// Library/Functions/Swap/SwapIecDate
FUNCTION SwapIecDate : IEC_DATE
// ------------------------------------------------------------------------- 
//  SRCI Robot Library                                                
// ------------------------------------------------------------------------- 
//                                                                           
//  Object:      SwapIecDate                                       
//  Author:      Thorsten Brach                                                
//  Date:        2024-06-09
//
//  Description:                                              
//   
//                                                                           
//  Copyright: 
//    (C) 2024 Thorsten Brach. All rights reserved                                                                                                                                            
//             Licensed under the MIT License.
//                                                                           
//  Disclaimer:                                                                           
//    This project is provided without any guarantee and can be used for   
//    private and commercial purposes. Any use is at the user’s 
//    own risk and responsibility.
//
// -------------------------------------------------------------------------
VAR_INPUT
  /// Value to swap
  Value : IEC_DATE;
END_VAR

SwapBytes(ADR(Value),SIZEOF(Value));

SwapIecDate := Value;

END_FUNCTION

// Library/Functions/Swap/SwapIecTime
FUNCTION SwapIecTime : TOD
// ------------------------------------------------------------------------- 
//  SRCI Robot Library                                                
// ------------------------------------------------------------------------- 
//                                                                           
//  Object:      SwapTime                                       
//  Author:      Thorsten Brach                                                
//  Date:        2024-06-01
//
//  Description:                                              
//   
//                                                                           
//  Copyright: 
//    (C) 2024 Thorsten Brach. All rights reserved                                                                                                                                            
//             Licensed under the MIT License.
//                                                                           
//  Disclaimer:                                                                           
//    This project is provided without any guarantee and can be used for   
//    private and commercial purposes. Any use is at the user’s 
//    own risk and responsibility.
//
// -------------------------------------------------------------------------
VAR_INPUT
  /// Value
  Value : TOD;
END_VAR

SwapBytes(ADR(Value),SIZEOF(Value));

SwapIecTime := Value;

END_FUNCTION

// Library/Functions/Swap/SwapInt
FUNCTION SwapInt : INT
// ------------------------------------------------------------------------- 
//  SRCI Robot Library                                                
// ------------------------------------------------------------------------- 
//                                                                           
//  Object:      SwapInt                                       
//  Author:      Thorsten Brach                                                
//  Date:        2024-06-01
//
//  Description:                                              
//   
//                                                                           
//  Copyright: 
//    (C) 2024 Thorsten Brach. All rights reserved                                                                                                                                            
//             Licensed under the MIT License.
//                                                                           
//  Disclaimer:                                                                           
//    This project is provided without any guarantee and can be used for   
//    private and commercial purposes. Any use is at the user’s 
//    own risk and responsibility.
//
// -------------------------------------------------------------------------
VAR_INPUT
  /// Value to swap
  Value : INT;
END_VAR

SwapBytes(ADR(Value),SIZEOF(Value));

SwapInt := Value;

END_FUNCTION

// Library/Functions/Swap/SwapReal
FUNCTION SwapReal : REAL
// ------------------------------------------------------------------------- 
//  SRCI Robot Library                                                
// ------------------------------------------------------------------------- 
//                                                                           
//  Object:      SwapReal                                       
//  Author:      Thorsten Brach                                                
//  Date:        2024-06-01
//
//  Description:                                              
//   
//                                                                           
//  Copyright: 
//    (C) 2024 Thorsten Brach. All rights reserved                                                                                                                                            
//             Licensed under the MIT License.
//                                                                           
//  Disclaimer:                                                                           
//    This project is provided without any guarantee and can be used for   
//    private and commercial purposes. Any use is at the user’s 
//    own risk and responsibility.
//
// -------------------------------------------------------------------------
VAR_INPUT
  /// Value
  Value : REAL;
END_VAR

SwapBytes(ADR(Value),SIZEOF(Value));

SwapReal := Value;

END_FUNCTION

// Library/Functions/Swap/SwapUdint
FUNCTION SwapUdint : UDINT
// ------------------------------------------------------------------------- 
//  SRCI Robot Library                                                
// ------------------------------------------------------------------------- 
//                                                                           
//  Object:      SwapUdint                                       
//  Author:      Thorsten Brach                                                
//  Date:        2024-06-01
//
//  Description:                                              
//   
//                                                                           
//  Copyright: 
//    (C) 2024 Thorsten Brach. All rights reserved                                                                                                                                            
//             Licensed under the MIT License.
//                                                                           
//  Disclaimer:                                                                           
//    This project is provided without any guarantee and can be used for   
//    private and commercial purposes. Any use is at the user’s 
//    own risk and responsibility.
//
// -------------------------------------------------------------------------
VAR_INPUT
  /// Value
  Value : UDINT;
END_VAR

SwapBytes(ADR(Value),SIZEOF(Value));

SwapUdint := Value;

END_FUNCTION

// Library/Functions/Swap/SwapUint
FUNCTION SwapUint : UINT
// ------------------------------------------------------------------------- 
//  SRCI Robot Library                                                
// ------------------------------------------------------------------------- 
//                                                                           
//  Object:      SwapUint                                       
//  Author:      Thorsten Brach                                                
//  Date:        2024-06-01
//
//  Description:                                              
//   
//                                                                           
//  Copyright: 
//    (C) 2024 Thorsten Brach. All rights reserved                                                                                                                                            
//             Licensed under the MIT License.
//                                                                           
//  Disclaimer:                                                                           
//    This project is provided without any guarantee and can be used for   
//    private and commercial purposes. Any use is at the user’s 
//    own risk and responsibility.
//
// -------------------------------------------------------------------------
VAR_INPUT
  /// Value to swap
  Value : UINT;
END_VAR

SwapBytes(ADR(Value),SIZEOF(Value));

SwapUint := Value;

END_FUNCTION

// Library/Interfaces/IMessageLogger
INTERFACE IMessageLogger

METHOD PUBLIC AddMessageLog
VAR_INPUT
  /// Message to add to the log
  MessageLog : AlarmMessage;
END_VAR
END_METHOD

METHOD PUBLIC AddSystemLog
VAR_INPUT
  /// System messafe to add to the log
  SystemLog : STRING(RobotLibraryParameter.MESSAGE_TEXT_LEN);
END_VAR
END_METHOD

END_INTERFACE

// Library/Interfaces/IRobotLibraryCommandFB
INTERFACE IRobotLibraryCommandFB

METHOD PUBLIC CallBack : DINT
VAR_INPUT
  /// Response data
  RspData : AxesGroupAcyclicAcrEntryRspBuffer;  
END_VAR
END_METHOD

PROPERTY CommandData : RobotLibrarySendDataFB
GET
END_GET
SET
END_SET
END_PROPERTY

END_INTERFACE

// Library/POUs/_internal/Send/RobotLibrarySendDataFB
{attribute 'pack_mode' := '1'} 
FUNCTION_BLOCK RobotLibrarySendDataFB extends RobotLibrarySendDataBaseFB
// ------------------------------------------------------------------------- 
//  SRCI Robot Library                                                
// ------------------------------------------------------------------------- 
//                                                                           
//  Object:      RobotLibrarySendDataFB                                      
//  Author:      Thorsten Brach                                                
//  Date:        2024-06-01
//
//  Description:                                              
//    
//                                                                           
//  Copyright: 
//    (C) 2024 Thorsten Brach. All rights reserved                                                                                                                                            
//             Licensed under the MIT License.
//                                                                           
//  Disclaimer:                                                                           
//    This project is provided without any guarantee and can be used for   
//    private and commercial purposes. Any use is at the user’s 
//    own risk and responsibility.
//
// -------------------------------------------------------------------------
VAR_INPUT
  /// Payload
  Payload     : POINTER TO BYTE;
  /// Size of the Payload array
  PayLoadSize : UDINT;
END_VAR

/// Resets the payload buffer, the payload pointer and the payload length
METHOD Reset
VAR_INPUT
END_VAR
SUPER^.Reset();

// Reset payload buffer
SysDepMemSet(pDest := Payload, Value := 0 , DataLen := PayLoadSize);
END_METHOD

METHOD SetLifeSignFooter
VAR_INPUT
  /// Life sign value
  LifeSign : BYTE;
END_VAR

VAR
  /// temporary 
  pLifeSign : POINTER TO BYTE;
END_VAR
pLifeSign := Payload + PayLoadSize -1;

pLifeSign^ := LifeSign;
END_METHOD

METHOD UpdatePointer
VAR_INPUT
END_VAR
pPayload := Payload;
END_METHOD

END_FUNCTION_BLOCK

// Library/POUs/_internal/Send/RobotLibrarySendDataBaseFB
{attribute 'pack_mode' := '1'} 
FUNCTION_BLOCK RobotLibrarySendDataBaseFB
// ------------------------------------------------------------------------- 
//  SRCI Robot Library                                                
// ------------------------------------------------------------------------- 
//                                                                           
//  Object:      RobotLibrarySendDataFB                                      
//  Author:      Thorsten Brach                                                
//  Date:        2024-06-01
//
//  Description:                                              
//    
//                                                                           
//  Copyright: 
//    (C) 2024 Thorsten Brach. All rights reserved                                                                                                                                            
//             Licensed under the MIT License.
//                                                                           
//  Disclaimer:                                                                           
//    This project is provided without any guarantee and can be used for   
//    private and commercial purposes. Any use is at the user’s 
//    own risk and responsibility.
//
// -------------------------------------------------------------------------
VAR_INPUT
  /// Payload length
  PayloadLen : UDINT;
  /// Payload pointer
  PayloadPtr : UDINT;
END_VAR


VAR
  /// internal pointer to payload 
  pPayload : POINTER TO BYTE;
END_VAR

/// Adds a ArmConfigParameter to the payload buffer, increase the payload pointer and returns the payload lenght
METHOD AddArmConfig : UDINT
VAR_INPUT
  /// Value to add
  Value : ArmConfigParameter;
END_VAR

VAR
  /// temporary Byte
 _tmpByte : BYTE;
END_VAR
// Table 6-274: "ConfigMode" on "Command Management Layer"
// --------------------------
// --------------------------
// Byte 00 : Bit 00  - Shoulder
//         : Bit 01  - Shoulder
//         : Bit 02  - Shoulder
//         : Bit 03  - Shoulder
//         : Bit 04  - Elbow
//         : Bit 05  - Elbow
//         : Bit 06  - Elbow
//         : Bit 07  - Elbow
// Byte 01 : Bit 00  - Wrist
//         : Bit 01  - Wrist
//         : Bit 02  - Wrist
//         : Bit 03  - Wrist
//         : Bit 04  - Reserve
//         : Bit 05  - Reserve
//         : Bit 06  - Reserve
//         : Bit 07  - Reserve
_tmpByte.0 := Value.Shoulder = ArmConfigShoulder.BACK;
_tmpByte.1 := Value.Elbow    = ArmConfigElbow.DOWN;
_tmpByte.2 := Value.Wrist    = ArmConfigWrist.FLIP;

AddByte(_tmpByte);
AddByte(0);

AddArmConfig := PayloadLen;
END_METHOD

/// Adds a BOOL to the payload buffer, increase the payload pointer and returns the payload lenght
METHOD AddBool : UDINT
VAR_INPUT
  /// Value to add
  Value : BOOL;
END_VAR

VAR
  /// temporary byte
 _tmpByte : BYTE := 0;
END_VAR
// update internal pointer
UpdatePointer();

// check pointer is valid ? 
IF (pPayload = RobotLibraryConstants.NULL_POINTER)
THEN
  RETURN;
END_IF


_tmpByte.0 := Value;
// copy data 
SysDepMemCpy(pDest := pPayload + PayloadPtr, pSrc := ADR(_tmpByte), DataLen := SIZEOF(_tmpByte));
// inc payload pointer 
PayloadPtr := PayloadPtr + SIZEOF(_tmpByte);
// return payload len
AddBool := PayloadLen := PayloadPtr;
END_METHOD

/// Adds a BYTE to the payload buffer, increase the payload pointer and returns the payload lenght
METHOD AddByte : UDINT
VAR_INPUT
  /// Value to add
  Value : BYTE;
END_VAR
// update internal pointer
UpdatePointer();

// check pointer is valid ? 
IF (pPayload = RobotLibraryConstants.NULL_POINTER)
THEN
  RETURN;
END_IF


Value := Value;
// copy data 
SysDepMemCpy( pDest := pPayload + PayloadPtr, pSrc := ADR(Value), DataLen := SIZEOF(Value));
// inc payload pointer 
PayloadPtr := PayloadPtr + SIZEOF(Value);
// return payload len
AddByte := PayloadLen := PayloadPtr;
END_METHOD

/// Adds a DataBlock to the payload buffer, increase the payload pointer and returns the payload lenght
METHOD AddDataBlock : UDINT
VAR_INPUT
  /// Value to add
  pValue : POINTER TO BYTE;
  /// Size of data block
  Size   : UDINT;
END_VAR
// update internal pointer
UpdatePointer();

// check pointer is valid ? 
IF (pPayload = RobotLibraryConstants.NULL_POINTER)
THEN
  RETURN;
END_IF


IF (pValue = 0) OR (Size = 0 )
THEN
  RETURN;
END_IF

// copy data 
SysDepMemCpy( pDest := pPayload + PayloadPtr, pSrc := pValue, DataLen := Size);
// inc payload pointer 
PayloadPtr := PayloadPtr + Size;
// return payload len
AddDataBlock := PayloadLen := PayloadPtr;
END_METHOD

/// Adds a DataInSync to the payload buffer, increase the payload pointer and returns the payload lenght
METHOD AddDataEnableSync : UDINT
VAR_INPUT
  /// Value to add
  Value : DataEnableSync;
END_VAR

VAR
  /// temporary Byte
 _tmpByte : BYTE;
END_VAR
Value := Value;

_tmpByte.0 := Value.EnableSyncTool;
_tmpByte.1 := Value.EnableSyncFrame;
_tmpByte.2 := Value.EnableSyncLoad;
_tmpByte.3 := Value.EnableSyncWorkArea;
_tmpByte.4 := Value.EnableSyncSWLimits;
_tmpByte.5 := Value.EnableSyncDefaultDynamics;
_tmpByte.6 := Value.EnableSyncReferenceDynamics;


AddByte(_tmpByte);

AddDataEnableSync := PayloadLen;
END_METHOD

/// Adds a DataInSync to the payload buffer, increase the payload pointer and returns the payload lenght
METHOD AddDataInSync : UDINT
VAR_INPUT
  /// Value to add
  Value : DataInSync;
END_VAR

VAR
  /// temporary Byte
 _tmpByte : BYTE;
END_VAR
Value := Value;

_tmpByte.0 := Value.ToolsInSync;
_tmpByte.1 := Value.FramesInSync;
_tmpByte.2 := Value.LoadsInSync;
_tmpByte.3 := Value.WorkAreasInSync;
_tmpByte.4 := Value.SoftwareLimitsInSync;
_tmpByte.5 := Value.DefaultDynamicsInSync;
_tmpByte.6 := Value.ReferenceDynamicsInSync;
_tmpByte.7 := FALSE;

AddByte(_tmpByte);

AddDataInSync := PayloadLen;
END_METHOD

/// Adds a DWORD to the payload buffer , increase the payload pointer and returns the payload lenght
METHOD AddDword : UDINT
VAR_INPUT
  /// Value to add
  Value : DWORD;
END_VAR
// update internal pointer
UpdatePointer();

// check pointer is valid ? 
IF (pPayload = RobotLibraryConstants.NULL_POINTER)
THEN
  RETURN;
END_IF


// swap byte order
Value := SwapDword(Value);
// copy data 
SysDepMemCpy(pDest := pPayload + PayloadPtr, pSrc := ADR(Value), DataLen := SIZEOF(Value));
// inc data index 
PayloadPtr := PayloadPtr + SIZEOF(Value);
// return payload len
AddDword := PayloadLen := PayloadPtr;
END_METHOD

/// Adds two halfe BYTE to the payload buffer , increase the payload pointer and returns the payload lenght
METHOD AddHalfBytes : UDINT
VAR_INPUT
  /// Value to add
  HalfByteHi : BYTE;
  /// Value to add
  HalfByteLo : BYTE;
END_VAR

VAR
  /// internal value
 _value : BYTE;
END_VAR
// update internal pointer
UpdatePointer();

// check pointer is valid ? 
IF (pPayload = RobotLibraryConstants.NULL_POINTER)
THEN
  RETURN;
END_IF


_value := CombineHalfBytes( HalfByteHi := HalfByteHi, HalfByteLo := HalfByteLo);
// copy data 
SysDepMemCpy(pDest := pPayload + PayloadPtr, pSrc := ADR(_value), DataLen := SIZEOF(_value));
// inc payload pointer 
PayloadPtr := PayloadPtr + SIZEOF(_value);
// return payload len
AddHalfBytes := PayloadLen := PayloadPtr;
END_METHOD

/// Adds a IEC_DATE to the payload buffer, increase the payload pointer and returns the payload lenght
METHOD AddIecDate : UDINT
VAR_INPUT
  /// Value to add
  Value : IEC_DATE;
END_VAR
// update internal pointer
UpdatePointer();

// check pointer is valid ? 
IF (pPayload = RobotLibraryConstants.NULL_POINTER)
THEN
  RETURN;
END_IF


Value := SwapIecDate(Value);
// copy data 
SysDepMemCpy(pDest := pPayload + PayloadPtr, pSrc := ADR(Value), DataLen := SIZEOF(Value));
// inc payload pointer 
PayloadPtr := PayloadPtr + SIZEOF(Value);
// return payload len
AddIecDate := PayloadLen := PayloadPtr;
END_METHOD

/// Adds a IEC_TIME to the payload buffer, increase the payload pointer and returns the payload lenght
METHOD AddIecTime : UDINT
VAR_INPUT
  /// Value to add
  Value : IEC_TIME;
END_VAR
// update internal pointer
UpdatePointer();

// check pointer is valid ? 
IF (pPayload = RobotLibraryConstants.NULL_POINTER)
THEN
  RETURN;
END_IF


Value := SwapIecTime(Value);
// copy data 
SysDepMemCpy(pDest := pPayload + PayloadPtr, pSrc := ADR(Value), DataLen := SIZEOF(Value));
// inc payload pointer 
PayloadPtr := PayloadPtr + SIZEOF(Value);
// return payload len
AddIecTime := PayloadLen := PayloadPtr;
END_METHOD

/// Adds a INT to the payload buffer , increase the payload pointer and returns the payload lenght
METHOD AddInt : UDINT
VAR_INPUT
  /// Value to add
  Value : INT;
END_VAR
// update internal pointer
UpdatePointer();

// check pointer is valid ? 
IF (pPayload = RobotLibraryConstants.NULL_POINTER)
THEN
  RETURN;
END_IF


// swap byte order
Value := SwapInt(Value);
// copy data 
SysDepMemCpy(pDest := pPayload + PayloadPtr, pSrc := ADR(Value), DataLen := SIZEOF(Value));
// inc data index 
PayloadPtr := PayloadPtr + SIZEOF(Value);
// return payload len
AddInt := PayloadLen := PayloadPtr;
END_METHOD

/// Adds a REAL to the payload buffer , increase the payload pointer and returns the payload lenght
METHOD AddReal : UDINT
VAR_INPUT
  /// Value to add
  Value : REAL;
END_VAR
// update internal pointer
UpdatePointer();

// check pointer is valid ? 
IF (pPayload = RobotLibraryConstants.NULL_POINTER)
THEN
  RETURN;
END_IF


// swap byte order
Value := SwapReal(Value);
// copy data 
SysDepMemCpy(pDest := pPayload + PayloadPtr,pSrc := ADR(Value), DataLen := SIZEOF(Value));
// inc data index 
PayloadPtr := PayloadPtr + SIZEOF(Value);
// return payload len
AddReal := PayloadLen := PayloadPtr;
END_METHOD

/// Adds a SINT to the payload buffer, increase the payload pointer and returns the payload lenght
METHOD AddSint : UDINT
VAR_INPUT
  /// Value to add
  Value : SINT;
END_VAR
// update internal pointer
UpdatePointer();

// check pointer is valid ? 
IF (pPayload = RobotLibraryConstants.NULL_POINTER)
THEN
  RETURN;
END_IF


Value := Value;
// copy data 
SysDepMemCpy(pDest := pPayload + PayloadPtr, pSrc := ADR(Value), DataLen := SIZEOF(Value));
// inc payload pointer 
PayloadPtr := PayloadPtr + SIZEOF(Value);
// return payload len
AddSint := PayloadLen := PayloadPtr;
END_METHOD

/// Adds a String to the payload buffer, increase the payload pointer and returns the payload lenght
METHOD AddString : UDINT
VAR_INPUT
  /// Value to add
  Value : STRING(255);
END_VAR
// update internal pointer
UpdatePointer();

// check pointer is valid ? 
IF (pPayload = RobotLibraryConstants.NULL_POINTER)
THEN
  RETURN;
END_IF


IF ( LEN(Value) = 0 )
THEN
  RETURN;
END_IF

// copy data 
SysDepMemCpy(pDest := pPayload + PayloadPtr, pSrc := ADR(Value), DataLen := DINT_TO_UDINT(LEN(Value)));
// inc payload pointer 
PayloadPtr := PayloadPtr + DINT_TO_UDINT(LEN(Value));
// return payload len
AddString := PayloadLen := PayloadPtr;
END_METHOD

/// Adds a TIME to the payload buffer , increase the payload pointer and returns the payload lenght
METHOD AddTime : UDINT
VAR_INPUT
  /// Value to add
  Value : TOD;
END_VAR
// update internal pointer
UpdatePointer();

// check pointer is valid ? 
IF (pPayload = RobotLibraryConstants.NULL_POINTER)
THEN
  RETURN;
END_IF


// swap byte order
Value := SwapIecTime(Value);
// copy data 
SysDepMemCpy(pDest := pPayload + PayloadPtr, pSrc := ADR(Value), DataLen := SIZEOF(Value));
// inc data index 
PayloadPtr := PayloadPtr + SIZEOF(Value);
// return payload len
AddTime := PayloadLen := PayloadPtr;
END_METHOD

/// Adds a TurnNumber to the payload buffer, increase the payload pointer and returns the payload lenght
METHOD AddTurnNumber : UDINT
VAR_INPUT
  /// Value to add
  Value : TurnNumber;
END_VAR

VAR
  /// temporary Byte
 _tmpByte : BYTE;
END_VAR
Value := Value;

// ST-FIX F3: sign + magnitude (spec 5.5.4.4)
AddHalfBytes( HalfByteHi := TURN_TO_SIGN_MAGNITUDE(Turns := Value.J2Turns, Bits := 3), HalfByteLo := TURN_TO_SIGN_MAGNITUDE(Turns := Value.J1Turns, Bits := 3));
AddHalfBytes( HalfByteHi := TURN_TO_SIGN_MAGNITUDE(Turns := Value.J4Turns, Bits := 3), HalfByteLo := TURN_TO_SIGN_MAGNITUDE(Turns := Value.J3Turns, Bits := 3));
AddHalfBytes( HalfByteHi := TURN_TO_SIGN_MAGNITUDE(Turns := Value.J6Turns, Bits := 3), HalfByteLo := TURN_TO_SIGN_MAGNITUDE(Turns := Value.J5Turns, Bits := 3));
AddByte(TURN_TO_SIGN_MAGNITUDE(Turns := Value.E1Turns, Bits := 7));

AddTurnNumber := PayloadLen;
END_METHOD

/// Adds a UDINT to the payload buffer , increase the payload pointer and returns the payload lenght
METHOD AddUdint : UDINT
VAR_INPUT
  /// Value to add
  Value : UDINT;
END_VAR
// update internal pointer
UpdatePointer();

// check pointer is valid ? 
IF (pPayload = RobotLibraryConstants.NULL_POINTER)
THEN
  RETURN;
END_IF


// swap byte order
Value := SwapUdint(Value);
// copy data 
SysDepMemCpy(pDest := pPayload + PayloadPtr, pSrc := ADR(Value), DataLen := SIZEOF(Value));
// inc data index 
PayloadPtr := PayloadPtr + SIZEOF(Value);
// return payload len
AddUdint := PayloadLen := PayloadPtr;
END_METHOD

/// Adds a UINT to the payload buffer , increase the payload pointer and returns the payload lenght
METHOD AddUint : UDINT
VAR_INPUT
  /// Value to add
  Value : UINT;
END_VAR
// update internal pointer
UpdatePointer();

// check pointer is valid ? 
IF (pPayload = RobotLibraryConstants.NULL_POINTER)
THEN
  RETURN;
END_IF


// swap byte order
Value := SwapUint(Value);
// copy data 
SysDepMemCpy(pDest := pPayload + PayloadPtr, pSrc := ADR(Value), DataLen := SIZEOF(Value));
// inc data index 
PayloadPtr := PayloadPtr + SIZEOF(Value);
// return payload len
AddUint := PayloadLen := PayloadPtr;
END_METHOD

/// Adds a USINT to the payload buffer, increase the payload pointer and returns the payload lenght
METHOD AddUsint : UDINT
VAR_INPUT
  /// Value to add
  Value : USINT;
END_VAR
// update internal pointer
UpdatePointer();

// check pointer is valid ? 
IF (pPayload = RobotLibraryConstants.NULL_POINTER)
THEN
  RETURN;
END_IF


Value := Value;
// copy data 
SysDepMemCpy(pDest := pPayload + PayloadPtr, pSrc := ADR(Value), DataLen := SIZEOF(Value));
// inc payload pointer 
PayloadPtr := PayloadPtr + SIZEOF(Value);
// return payload len
AddUsint := PayloadLen := PayloadPtr;
END_METHOD

/// Resets the payload buffer, the payload pointer and the payload length
METHOD Reset
VAR_INPUT
END_VAR
PayloadLen := 0;
PayloadPtr := 0;
END_METHOD

METHOD UpdatePointer
VAR_INPUT
END_VAR
END_METHOD

END_FUNCTION_BLOCK

// Library/POUs/_internal/BaseFBs/RobotLibraryBaseEnableFB
FUNCTION_BLOCK RobotLibraryBaseEnableFB EXTENDS RobotLibraryBaseFB
// ------------------------------------------------------------------------- 
//  SRCI Robot Library                                                
// ------------------------------------------------------------------------- 
//                                                                           
//  Object:      RobotLibraryBaseFB                                       
//  Author:      Thorsten Brach                                                
//  Date:        2024-08-11
//
//  Description:                                              
//   
//                                                                           
//  Copyright: 
//    (C) 2024 Thorsten Brach. All rights reserved                                                                                                                                            
//             Licensed under the MIT License.
//                                                                           
//  Disclaimer:                                                                           
//    This project is provided without any guarantee and can be used for   
//    private and commercial purposes. Any use is at the user’s 
//    own risk and responsibility.
//
// -------------------------------------------------------------------------
VAR_INPUT
  /// Set TRUE to activate / Set False to deactivate
  Enable            : BOOL;
END_VAR

VAR_OUTPUT
  /// FB is being processed
  Busy              : BOOL;
  /// TRUE while function is active
  Enabled           : BOOL;
END_VAR

VAR
  /// Rising edge for enable
  {attribute 'hide'}
 _enable_R          : R_TRIG;
  /// Falling edge for enable
  {attribute 'hide'}
 _enable_F          : F_TRIG;
END_VAR

SUPER^(AxesGroup := AxesGroup);

// ST-FIX F135: "Enabled" is reset with the falling edge of "Enable" as soon as possible
// (spec 5.5.10 output status), also while the FB still sends the deactivation to the RC
IF ( NOT Enable )
THEN
  Enabled := FALSE;
END_IF

METHOD PROTECTED OnCall
VAR_IN_OUT
  /// Robot assignment of function
  AxesGroup : AxesGroup; 
END_VAR

VAR
  /// internal return value
 _retVal : DINT;
END_VAR

                  SUPER^.OnCall(AxesGroup := AxesGroup);

// building rising and falling edges
_enable_R( CLK := Enable);
_enable_F( CLK := Enable);


// Check command execution is allowed ?
IF ((     Enable                                 ) AND
    ( NOT AxesGroup.State.Initialized            ) AND
    ( NOT AxesGroup.State.Synchronized           ) AND
    (     MyType <> 'MC_ExchangeConfigurationFB' ) AND // is part of init sequence
    (     MyType <> 'MC_ReadMessagesFB'          ) AND // is part of init sequence
    (     MyType <> 'MC_ReadRobotDataFB'         ))    // is part of init sequence
THEN
  SetError( ErrorID := RobotLibraryErrorIdEnum.ERR_COMMANDS_NOT_ENABLED, Overwrite := TRUE );
  Error   := TRUE;
  Busy    := FALSE; 
END_IF


// On execution started
IF ( _enable_R.Q )
THEN
  // ST-FIX F23: a new enable ends a pending cancel / error clear of the previous enable
  _cancel := FALSE;
  _stepCancel := 0;
  _clearError := FALSE;
  _stepClearError := 0;
  // ST-FIX F78: an error of the previous enable that is still being cleared (falling edge, up
  // to 5 s) is cleared now - otherwise the block (start only without Error) consumes the
  // rising edge and the new enable is ignored (not sent, no Busy, no Error)
  IF ( Error ) AND ( ErrorID <> RobotLibraryErrorIdEnum.ERR_COMMANDS_NOT_ENABLED )
  THEN
    Reset();
  END_IF
  OnExecStart(AxesGroup := AxesGroup);
END_IF


// On execution cancel  
IF ( Busy ) AND ( _enable_F.Q ) 
THEN
  // set cancel flag
 _cancel := TRUE;
END_IF

IF ( _cancel )
THEN
  // call Cancel
 _retVal := OnExecCancel(AxesGroup := AxesGroup);
  
  // done or error ?
  IF ( _retVal <> RobotLibraryConstants.RUNNING )
  THEN
    // reset cancel flag
   _cancel := FALSE;
	END_IF
END_IF


// On execution error clear
IF ( Error ) AND ( _enable_F.Q )
THEN
  // set ClearError flag
 _clearError := TRUE;
END_IF

IF ( _clearError )
THEN
 _retVal := OnExecErrorClear(AxesGroup := AxesGroup); 

  // done or error ?
  IF ( _retVal <> RobotLibraryConstants.RUNNING )
  THEN
    // reset ClearError flag
   _clearError := FALSE;
	END_IF
END_IF
END_METHOD

METHOD Protected OnExecCancel : DINT
VAR_IN_OUT
  /// Robot assignment of function
  AxesGroup : AxesGroup; 
END_VAR
VAR
  /// internal return value 
 _retVal    : DINT;
END_VAR
OnExecCancel := Reset();

// Create log entry
CreateLogMessagePara1 ( Timestamp   := AxesGroup.State.SystemTime,
                        MessageType := MessageType.CMD,
                        Severity    := Severity.DEBUG,
                        MessageCode := 0,
                        MessageText := 'Execution of {1} cancled ',
                        Para1       := MyType);                 

// try to remove cmd
_retVal := AxesGroup.Acyclic.ActiveCommandRegister.RemoveCmd(_uniqueID);

IF (_retVal = RobotLibraryConstants.OK)
THEN
  // Create log entry
  CreateLogMessagePara1 ( Timestamp   := AxesGroup.State.SystemTime,
                          MessageType := MessageType.CMD,
                          Severity    := Severity.DEBUG,
                          MessageCode := 0,
                          MessageText := '{1} successfully removed from ACR',
                          Para1       := MyType);                 
ELSE
  // Create log entry
  CreateLogMessagePara1 ( Timestamp   := AxesGroup.State.SystemTime,
                          MessageType := MessageType.CMD,
                          Severity    := Severity.DEBUG,
                          MessageCode := 0,
                          MessageText := '{1} was not removed from ACR because execution was already in progress',
                          Para1       := MyType);                 
END_IF
END_METHOD

METHOD PROTECTED OnExecErrorClear : DINT
VAR_IN_OUT
  /// Robot assignment of function
  AxesGroup : AxesGroup; 
END_VAR
OnExecErrorClear := RobotLibraryConstants.RUNNING;

CASE _stepClearError OF
  
  0:  // Reset 
      Reset();
      // trigger parameter update to disable FB
     _parameterUpdateInternal := TRUE;
      // call Check Parameter changed method to trigger the parameter update to deactivate jogging mode
      CheckParameterChanged(AxesGroup := AxesGroup);
      // set timeout
      SetTimeout(PT := _timeoutClearError, rTimer := _timerClearError);
      // inc step counter
     _stepClearError := _stepClearError + 1; 
      
  1: IF ( _responseReceived )
     THEN     
       // reset response received flag
      _responseReceived := FALSE;
       // reset step counter
      _stepClearError := 0;
       // finished
       OnExecErrorClear := RobotLibraryConstants.OK;
     ELSE
       // timeout exceeded ? 
       IF (CheckTimeout(_timerClearError) = RobotLibraryConstants.OK)
       THEN
         OnExecErrorClear := RobotLibraryConstants.HAS_ERROR;
       END_IF
	   END_IF
ELSE
  // invalid step
  SetError( ErrorID := RobotLibraryErrorIdEnum.ERR_INVALID_STEP, Overwrite := TRUE );
END_CASE


// reset step counter
IF (OnExecErrorClear <> RobotLibraryConstants.RUNNING)
THEN
 _stepClearError := 0;
END_IF
END_METHOD

METHOD PROTECTED OnExecRun : DINT
VAR_IN_OUT
  /// Robot assignment of function
  AxesGroup : AxesGroup; 
END_VAR
END_METHOD

METHOD PROTECTED OnExecStart : DINT
VAR_IN_OUT
  /// Robot assignment of function
  AxesGroup : AxesGroup; 
END_VAR


// ST-FIX F71: Priority (1 = very high ... 4 = low, table 7-1)
IF ( Priority < PriorityLevel.VERY_HIGH )
THEN
  SetError( ErrorID := RobotLibraryErrorIdEnum.ERR_PRIORITY_TOO_HIGH, Overwrite := TRUE );
  // Create log entry
  CreateLogMessage ( Timestamp   := AxesGroup.State.SystemTime,
                     MessageType := MessageType.CMD,
                     Severity    := Severity.ERROR,
                     MessageCode := ErrorID,
                     MessageText := 'Invalid input Priority: higher than VERY_HIGH');
  Error := TRUE;
ELSIF ( Priority > PriorityLevel.LOW )
THEN
  SetError( ErrorID := RobotLibraryErrorIdEnum.ERR_PRIORITY_TOO_LOW, Overwrite := TRUE );
  // Create log entry
  CreateLogMessage ( Timestamp   := AxesGroup.State.SystemTime,
                     MessageType := MessageType.CMD,
                     Severity    := Severity.ERROR,
                     MessageCode := ErrorID,
                     MessageText := 'Invalid input Priority: lower than LOW');
  Error := TRUE;
END_IF
END_METHOD

METHOD PROTECTED OnUpdateStateFlags
VAR_INPUT
  /// Command message state
  State : CmdMessageState;
END_VAR
CASE State OF

  // No operation or process is active
  CmdMessageState.EMPTY               :;
  // Created but not yet started
  CmdMessageState.CREATED             :;
  // Buffered and awaiting execution
  CmdMessageState.BUFFERED            :;
  // Buffered in planner for future execution
  CmdMessageState.BUFFERED_IN_PLANNER :;
  // Currently active and in progress
  CmdMessageState.ACTIVE              :;
  // Interrupted and awaiting continuation
  CmdMessageState.INTERRUPTED         :;
  // Requested for abort
  CmdMessageState.ABORT_REQUEST       :;
  // Successfully completed
  CmdMessageState.DONE                : Busy := FALSE;
  // Aborted before completion
  CmdMessageState.ABORTED             : Busy := FALSE;
  // Encountered an error during execution
  CmdMessageState.ERROR               : Busy := FALSE;
END_CASE
END_METHOD

METHOD PROTECTED Reset : DINT
VAR_INPUT
END_VAR
Reset := SUPER^.Reset();

Busy    := FALSE;
Enabled := FALSE;
END_METHOD

END_FUNCTION_BLOCK

// Library/POUs/_internal/BaseFBs/RobotLibraryBaseFB

            
              FUNCTION_BLOCK RobotLibraryBaseFB EXTENDS RobotLibraryLogFB
// ------------------------------------------------------------------------- 
//  SRCI Robot Library                                                
// ------------------------------------------------------------------------- 
//                                                                           
//  Object:      RobotLibraryBaseFB                                       
//  Author:      Thorsten Brach                                                
//  Date:        2024-06-01
//
//  Description:                                              
//   
//                                                                           
//  Copyright: 
//    (C) 2024 Thorsten Brach. All rights reserved                                                                                                                                            
//             Licensed under the MIT License.
//                                                                           
//  Disclaimer:                                                                           
//    This project is provided without any guarantee and can be used for   
//    private and commercial purposes. Any use is at the user’s 
//    own risk and responsibility.
//
// -------------------------------------------------------------------------
VAR_INPUT
  /// User defined command name
  Name         : STRING(80);
  /// Execution Mode
  ExecMode     : ExecutionMode;
  /// Priority
  Priority     : PriorityLevel;
END_VAR
VAR_OUTPUT
  /// Command data
  CommandData  : RobotLibraryCommandDataFB;
  /// response data
  ResponseData : RobotLibraryResponseDataFB;
  /// An error occurred during the execution of the command
  Error        : BOOL;
  /// ErrorID reported by RC for error identification according to Table 7-1
  ErrorID      : WORD;
  ErrorIdEnum  : RobotLibraryErrorIdEnum;  
  ErrorAddTxt  : STRING(RobotLibraryConstants.MAX_ADD_TEXT_LENGTH);
  
  /// WarningID for warning identification reported during execution of command according to Table 7-3
  WarningID    : WORD;
  WarningIdEnum: RobotLibraryWarningIdEnum;  
  /// InfoID for info identification reported during execution of command according to Table 7-5
  InfoID       : WORD;    
  InfoIdEnum   : RobotLibraryInfoIdEnum;  
END_VAR
VAR_IN_OUT
  /// Robot assignment of function
  AxesGroup    : AxesGroup; 
END_VAR

VAR
  /// Rising edge for error
  {attribute 'hide'}
 _error_R                  : R_TRIG;
  /// Rising edge for warning
  {attribute 'hide'}
 _warning_R                : R_TRIG;
  /// Rising edge for information
  {attribute 'hide'}
 _info_R                   : R_TRIG;
  /// clear error active
 _clearError               : BOOL;
  /// cancel active
 _cancel                   : BOOL; 
  /// unique ID
 _uniqueID                 : UDINT;  
  /// flag for response received
 _responseReceived         : BOOL;
  /// internal step counter
 _stepCmd                  : DINT;
  /// internal timer  
  {attribute 'hide'}
 _timerCmd                 : TON;
  /// internal timeout 
  {attribute 'hide'}
 _timeoutCmd               : TIME := T#5S;
  /// internal step counter for ClearError
 _stepClearError           : DINT;
  /// internal timer for ClearError
  {attribute 'hide'}
 _timerClearError          : TON;
  /// internal timeout for ClearError 
  {attribute 'hide'}
 _timeoutClearError        : TIME := T#5S;

  /// internal step counter for Cancel
 _stepCancel               : DINT;
  /// internal timer for Cancel  
  {attribute 'hide'}
 _timerCancel              : TON;
  /// internal timeout for Cancel 
  {attribute 'hide'}
 _timeoutCancel            : TIME := T#5S;

  /// internal command header
 _cmdHeader                : CmdHeader;  
  /// internal response header
 _rspHeader                : RspHeader;
  /// internal flag for send a parameter update
 _parameterUpdateInternal  : BOOL; 
  /// internal flag for parameter has changed
 _parameterChanged         : BOOL;
  /// internal flag for parameter are valid
 _parameterValid           : BOOL;
END_VAR
            
          
VAR
  /// ST-FIX F74: message of the command for the message buffer
  _alarmMessage : AlarmMessage;
END_VAR
VAR
  /// ST-FIX F105: block type and command name for the messages
  _messageSource : STRING;
END_VAR

            
          
VAR
  /// ST-FIX F116: axes group of the running command
  _axesGroupAdr    : POINTER TO AxesGroup;
  /// ST-FIX F116: _axesGroupAdr is valid
  _axesGroupStored : BOOL;
END_VAR


            
            // ST-FIX F116: the AxesGroup input must not change while a command of this block is running
  IF ( _uniqueID <> 0 ) AND ( _axesGroupStored ) AND ( NOT Error )
  THEN
    IF ( _axesGroupAdr <> ADR(AxesGroup) )
    THEN
      _axesGroupAdr^.Acyclic.ActiveCommandRegister.RemoveCmd( UniqueID := _uniqueID );
      SetError( ErrorID := RobotLibraryErrorIdEnum.ERR_AXESGROUP_CHANGED, Overwrite := TRUE );
      // Create log entry (the command keeps running on the RC of the first axes group)
      CreateLogMessagePara1 ( Timestamp   := AxesGroup.State.SystemTime,
                              MessageType := MessageType.CMD,
                              Severity    := Severity.ERROR,
                              MessageCode := ErrorID,
                              MessageText := 'AxesGroup of {1} changed while the command was running',
                              Para1       := MyType);
      OnUpdateStateFlags( State := CmdMessageState.ERROR );
    END_IF
  END_IF
  IF ( _uniqueID = 0 )
  THEN
    _axesGroupStored := FALSE;
  ELSIF ( NOT _axesGroupStored )
  THEN
    _axesGroupAdr    := ADR(AxesGroup);
    _axesGroupStored := TRUE;
  END_IF

  OnCall               (AxesGroup := AxesGroup);
OnExecRun            (AxesGroup := AxesGroup);
// ST-FIX F53: no response of the RC within _timeoutCmd after the command was added
// -> error (before: _timerCmd was started but never evaluated, the FB stayed Busy)
IF ( _uniqueID <> 0 ) AND ( _rspHeader.State = CmdMessageState.EMPTY ) AND ( NOT Error )
THEN
  IF ( CheckTimeout( rTimer := _timerCmd ) = RobotLibraryConstants.OK )
  THEN
    AxesGroup.Acyclic.ActiveCommandRegister.RemoveCmd( UniqueID := _uniqueID );
    SetError( ErrorID := RobotLibraryErrorIdEnum.ERR_TIMEOUT_CMD, Overwrite := TRUE );
    // Create log entry
    CreateLogMessage ( Timestamp   := AxesGroup.State.SystemTime,
                       MessageType := MessageType.CMD,
                       Severity    := Severity.ERROR,
                       MessageCode := ErrorID,
                       MessageText := 'No response of the RC within the command timeout');
    OnUpdateStateFlags( State := CmdMessageState.ERROR );
  END_IF
END_IF
CheckParameterChanged(AxesGroup := AxesGroup);


IF ( AxesGroup.State.OnlineChange_R.Q )
THEN
  OnOnlineChange(AxesGroup := AxesGroup);
END_IF
// ST-FIX F61: Error follows ErrorID in the same cycle, and with Error the other state outputs
// are reset (Busy/Active/Done/CommandAborted exclusive, spec table 5-45)
Error := ErrorID <> RobotLibraryConstants.OK;
IF ( Error )
THEN
  OnUpdateStateFlags( State := CmdMessageState.ERROR );
END_IF

METHOD PUBLIC CallBack : DINT
VAR_INPUT
  /// Response data
  RspData   : AxesGroupAcyclicAcrEntryRspBuffer;  
  /// Timestamp
  Timestamp : SystemTime;
END_VAR
// Create log entry
CreateLogMessagePara2 ( Timestamp   := Timestamp,
                        MessageType := MessageType.CMD,
                        Severity    := Severity.DEBUG,
                        MessageCode := 0,
                        MessageText := 'Callback reveiced in FB {1} <{2}>',
                        Para1       := MyType,
                        Para2       := Name);

                   
                   
ResponseData.Reset();
ResponseData.Payload    := RspData.Payload; 
ResponseData.PayloadLen := RspData.PayloadLen;
ParseResponsePayload( ResponseData :=  ResponseData , Timestamp := Timestamp);

// set flag for response received
_responseReceived := TRUE;
// ST-FIX F61: Error follows ErrorID in the same cycle, and with Error the other state outputs
// are reset (Busy/Active/Done/CommandAborted exclusive, spec table 5-45)
Error := ErrorID <> RobotLibraryConstants.OK;
IF ( Error )
THEN
  OnUpdateStateFlags( State := CmdMessageState.ERROR );
END_IF
END_METHOD

METHOD PROTECTED CheckFunctionSupported : BOOL
VAR_IN_OUT
  /// Robot assignment of function
  AxesGroup : AxesGroup; 
END_VAR
Error       := TRUE;
ErrorID     := RobotLibraryErrorIdEnum.ERR_FUNCTION_NOT_SUPPORTED;
ErrorAddTxt := CONCAT(THIS^._myType, ' ');
ErrorAddTxt := CONCAT(ErrorAddTxt , THIS^.Name);


// Create log entry
CreateLogMessagePara1 ( Timestamp   := AxesGroup.State.SystemTime,
                        MessageType := MessageType.CMD,
                        Severity    := Severity.DEBUG,
                        MessageCode := 0,
                        MessageText := 'Execution canceled, because function <{1}> is not supported by the robot controller',
                        Para1       :=  _myType);
END_METHOD

METHOD PROTECTED CheckParameterChanged : BOOL
VAR_IN_OUT
  /// Robot assignment of function
  AxesGroup    : AxesGroup; 
END_VAR
IF ( CheckParameterChanged )
THEN
  AxesGroup.Acyclic.ActiveCommandRegister.NotifyParameterChanged := _uniqueID;
END_IF
END_METHOD

METHOD PROTECTED CheckParameterValid : BOOL
VAR_IN_OUT
  /// Robot assignment of function
  AxesGroup : AxesGroup; 
END_VAR
CheckParameterValid := TRUE;
END_METHOD

METHOD INTERNAL CreateCommandPayload : RobotLibraryCommandDataFB
VAR_IN_OUT
  /// Robot assignment of function
  AxesGroup    : AxesGroup; 
END_VAR
// Reset all variables
CreateCommandPayload.Reset();
// Add CmdType
CreateCommandPayload.AddUint(_cmdHeader.CmdTyp);
// Add Reserve_ExecMode
CreateCommandPayload.AddHalfBytes(  0               , _cmdHeader.ExecMode);
// Add ParSeq_Priority
CreateCommandPayload.AddHalfBytes( _cmdHeader.ParSeq, _cmdHeader.Priority);

// ST-FIX F48: undefined ExecutionMode (spec table 5-75) -> error, not sent
CASE _cmdHeader.ExecMode OF
  ExecutionMode.SEQUENCE_PRIMARY, ExecutionMode.SEQUENCE_ABORT_OTHERS_PRIMARY,
  ExecutionMode.PARALLEL, ExecutionMode.CONTINUOUS, ExecutionMode.TRIGGER_MULTIPLE,
  ExecutionMode.SEQUENCE_SECONDARY, ExecutionMode.SEQUENCE_ABORT_OTHERS_SECONDARY,
  ExecutionMode.STOP_PARALLEL_CONTINUOUS_TRIGGER: ;
ELSE
  SetError( ErrorID := RobotLibraryErrorIdEnum.ERR_INVALID_PARAM_EXECUTION_MODE, Overwrite := TRUE );
  // Create log entry
  CreateLogMessagePara1 ( Timestamp   := AxesGroup.State.SystemTime,
                          MessageType := MessageType.CMD,
                          Severity    := Severity.ERROR,
                          MessageCode := ErrorID,
                          MessageText := 'Invalid ExecutionMode = {1}',
                          Para1       := EXECUTION_MODE_TO_STRING(_cmdHeader.ExecMode));
  OnUpdateStateFlags( State := CmdMessageState.ERROR );
END_CASE
END_METHOD

PROPERTY PUBLIC HasError : Bool
GET
HasError := ErrorID <> RobotLibraryErrorIdEnum.NO_ERROR;
END_GET
END_PROPERTY

PROPERTY PUBLIC HasInfo : BOOL
GET
HasInfo := InfoID <> RobotLibraryInfoIdEnum.NO_INFO;
END_GET
END_PROPERTY

PROPERTY PUBLIC HasWarning : BOOL
GET
HasWarning := WarningID <> RobotLibraryWarningIdEnum.NO_WARNING;
END_GET
END_PROPERTY

METHOD PROTECTED OnApplyOutCmd
VAR_INPUT
  /// Command message state
  State : CmdMessageState;
END_VAR
END_METHOD

METHOD PROTECTED OnCall
VAR_IN_OUT
  /// Robot assignment of function
  AxesGroup : AxesGroup; 
END_VAR
// map numeric value to enum, so that the corresponding message text is directly shown by the tooltip
ErrorIdEnum   := ErrorId;
WarningIdEnum := WarningId;
InfoIdEnum    := InfoId;

Error := ErrorID <> RobotLibraryConstants.OK;

InternalLogger   := AxesGroup.MessageLog; 
ExternalLogger   := AxesGroup.MessageLog.ExternalLogger;
LogLevel         := AxesGroup.MessageLog.LogLevel;

// building rising edges for error, warning, info number detected
_error_R  ( CLK := ErrorID   <> RobotLibraryConstants.OK );
_warning_R( CLK := WarningID <> RobotLibraryConstants.OK );
_info_R   ( CLK := InfoID    <> RobotLibraryConstants.OK );


// ST-FIX F105: the user defined command name belongs into the message text (spec 5.5.11,
// table 5-47 "[Robot] [Client] [MoveLinAbs] [MoveToP1] [text]")
_messageSource := MyType;
IF ( Name <> '' )
THEN
  _messageSource := CONCAT(MyType, CONCAT(' [', CONCAT(Name, ']')));
END_IF

// ST-FIX F74: every message of the command - also the client-side ones (e.g. parameter errors,
// before: only with the severity of the last response of the RC) - goes into the message
// buffer, with ACR entry and command type
IF ( _error_R.Q ) AND ( LogLevel <= Severity.ERROR ) (* ST-FIX F164: was < *)
THEN
  _alarmMessage.Severity    := Severity.ERROR;
  IF ( ErrorID = _rspHeader.AlarmMessageCode ) AND ( _rspHeader.AlarmMessageSeverity > Severity.ERROR )
  THEN
    _alarmMessage.Severity  := _rspHeader.AlarmMessageSeverity; // e.g. fatal error of the RC
  END_IF
  _alarmMessage.Timestamp   := AxesGroup.State.SystemTime;
  _alarmMessage.MessageType := MessageType.CMD;
  _alarmMessage.MessageCode := ErrorID;
  _alarmMessage.AcrID       := UDINT_TO_UINT(_uniqueID);
  _alarmMessage.CmdType     := _cmdHeader.CmdTyp;
  _alarmMessage.MessageText := CONCAT(_messageSource, CONCAT(' : ', MESSAGE_CODE_TO_STRING(ErrorID))); // ST-FIX F105
  AxesGroup.MessageLog.AddMessageLog( MessageLog := _alarmMessage );
END_IF
IF ( _warning_R.Q ) AND ( LogLevel <= Severity.WARNING ) (* ST-FIX F164: was < *)
THEN
  _alarmMessage.Severity    := Severity.WARNING;
  IF ( WarningID = _rspHeader.AlarmMessageCode ) AND ( _rspHeader.AlarmMessageSeverity > Severity.WARNING )
  THEN
    _alarmMessage.Severity  := _rspHeader.AlarmMessageSeverity; // e.g. fatal error of the RC
  END_IF
  _alarmMessage.Timestamp   := AxesGroup.State.SystemTime;
  _alarmMessage.MessageType := MessageType.CMD;
  _alarmMessage.MessageCode := WarningID;
  _alarmMessage.AcrID       := UDINT_TO_UINT(_uniqueID);
  _alarmMessage.CmdType     := _cmdHeader.CmdTyp;
  _alarmMessage.MessageText := CONCAT(_messageSource, CONCAT(' : ', MESSAGE_CODE_TO_STRING(WarningID))); // ST-FIX F105
  AxesGroup.MessageLog.AddMessageLog( MessageLog := _alarmMessage );
END_IF
IF ( _info_R.Q ) AND ( LogLevel <= Severity.INFO ) (* ST-FIX F164: was < *)
THEN
  _alarmMessage.Severity    := Severity.INFO;
  IF ( InfoID = _rspHeader.AlarmMessageCode ) AND ( _rspHeader.AlarmMessageSeverity > Severity.INFO )
  THEN
    _alarmMessage.Severity  := _rspHeader.AlarmMessageSeverity; // e.g. fatal error of the RC
  END_IF
  _alarmMessage.Timestamp   := AxesGroup.State.SystemTime;
  _alarmMessage.MessageType := MessageType.CMD;
  _alarmMessage.MessageCode := InfoID;
  _alarmMessage.AcrID       := UDINT_TO_UINT(_uniqueID);
  _alarmMessage.CmdType     := _cmdHeader.CmdTyp;
  _alarmMessage.MessageText := CONCAT(_messageSource, CONCAT(' : ', MESSAGE_CODE_TO_STRING(InfoID))); // ST-FIX F105
  AxesGroup.MessageLog.AddMessageLog( MessageLog := _alarmMessage );
END_IF
 


IF ( _error_R.Q)
THEN
  // Create log entry
  CreateLogMessagePara2 ( Timestamp   := AxesGroup.State.SystemTime,
                          MessageType := MessageType.CMD,
                          Severity    := Severity.DEBUG,
                          MessageCode := 0,
                          MessageText := 'Error with ID: 16#{1} in FB {2} received ',
                          Para1       := WORD_TO_STRING_HEX(ErrorID),
                          Para2       := MyType);                        
END_IF

IF ( _warning_R.Q)
THEN
  // Create log entry
  CreateLogMessagePara2 ( Timestamp   := AxesGroup.State.SystemTime,
                          MessageType := MessageType.CMD,
                          Severity    := Severity.DEBUG,
                          MessageCode := 0,
                          MessageText := 'Warning with ID: 16#{1} in FB {2} received ',
                          Para1       := WORD_TO_STRING_HEX(WarningID),
                          Para2       := MyType);                        
END_IF

IF ( _info_R.Q)
THEN
  // Create log entry
  CreateLogMessagePara2 ( Timestamp   := AxesGroup.State.SystemTime,
                          MessageType := MessageType.CMD,
                          Severity    := Severity.DEBUG,
                          MessageCode := 0,
                          MessageText := 'Info with ID: 16#{1} in FB {2} received ',
                          Para1       := WORD_TO_STRING_HEX(InfoID),
                          Para2       := MyType);                        
END_IF
END_METHOD

METHOD PROTECTED OnExecRun : DINT
VAR_IN_OUT
  /// Robot assignment of function
  AxesGroup : AxesGroup; 
END_VAR
END_METHOD

METHOD OnOnlineChange : DINT
VAR_IN_OUT
  /// Robot assignment of function
  AxesGroup : AxesGroup; 
END_VAR
// update pointer to command FB
AxesGroup.Acyclic.ActiveCommandRegister.OnOnlineChange( UniqueID := _uniqueID, pCommandFB := ADR(THIS^));
END_METHOD

METHOD PROTECTED OnUpdateStateFlags
VAR_INPUT
  /// Command message state
  State : CmdMessageState;
END_VAR
END_METHOD

METHOD INTERNAL ParseResponsePayload : DINT
VAR_INPUT
  /// Response data
  ResponseData : RobotLibraryResponseDataFB;
  /// Timestamp
  Timestamp    : SystemTime;  
END_VAR
// reset message IDs 
// ST-FIX F62: InfoID/WarningID/ErrorID are held until the falling edge of Execute/Enable
// (Reset), a response without message must not clear them (spec 5.5.10)

// get State
_rspHeader.State                := ResponseData.GetHalfeByte1(IncPayloadPtr := FALSE);
// get ParSeq
_rspHeader.ParSeq               := ResponseData.GetHalfeByte2(IncPayloadPtr := TRUE);
// get AlarmMessageSeverity
_rspHeader.AlarmMessageSeverity := ResponseData.GetSint();
// get AlarmMessageCode
_rspHeader.AlarmMessageCode     := ResponseData.GetUint();


// Update InfoID / WarningID / ErrorID
CASE _rspHeader.AlarmMessageSeverity OF

  // Informative message
  Severity.INFO        : SetInfo   ( InfoID    := _rspHeader.AlarmMessageCode, Overwrite := TRUE );
  // Warning message
  Severity.WARNING     : SetWarning( WarningID := _rspHeader.AlarmMessageCode, Overwrite := TRUE );
  // Error message
  Severity.ERROR       : SetError  ( ErrorID   := _rspHeader.AlarmMessageCode, Overwrite := TRUE ); 
  // Fataö error message
  Severity.FATAL_ERROR : SetError  ( ErrorID   := _rspHeader.AlarmMessageCode, Overwrite := TRUE );

END_CASE

// ST-FIX F61: state ERROR without error code (or with severity INFO/WARNING) -> 16#8613
IF ( _rspHeader.State = CmdMessageState.ERROR ) AND ( ErrorID = RobotLibraryConstants.OK )
THEN
  SetError( ErrorID := RobotLibraryErrorIdEnum.ERR_ROBOT_ERROR_NO_ID, Overwrite := TRUE );
  // Create log entry
  CreateLogMessage ( Timestamp   := Timestamp,
                     MessageType := MessageType.CMD,
                     Severity    := Severity.ERROR,
                     MessageCode := ErrorID,
                     MessageText := 'Response of the RC with state ERROR but without error code');
END_IF
ParseResponsePayload := ResponseData.PayloadPtr;
END_METHOD

METHOD PROTECTED Reset : DINT
VAR_INPUT
END_VAR
_parameterUpdateInternal := FALSE;
_responseReceived := FALSE;

_uniqueId := 0;
_rspHeader.State := CmdMessageState.EMPTY; // ST-FIX F53: no response yet
_stepCmd  := 0;
Error     := FALSE;
ErrorID   := 0;
WarningID := 0;
InfoID    := 0;  

Reset := RobotLibraryConstants.OK;
END_METHOD

METHOD PUBLIC SetError
VAR_INPUT
  /// ErrorID reported by RC for error identification according to Table 7-1
  ErrorID   : WORD;
  /// TRUE = overwrite an existing error 
  Overwrite : BOOL;
END_VAR
IF ( NOT HasError ) OR ( Overwrite )
THEN
  THIS^.ErrorID := ErrorID;
END_IF
END_METHOD

METHOD PUBLIC SetInfo
VAR_INPUT
  /// InfoID for info identification reported during execution of command according to Table 7-5
  InfoID    : WORD;
  /// TRUE = overwrite an existing info 
  Overwrite : BOOL;
END_VAR
IF ( NOT HasInfo ) OR ( Overwrite )
THEN
  THIS^.InfoID := InfoID;
END_IF
END_METHOD

METHOD PUBLIC SetWarning
VAR_INPUT
  /// WarningID for warning identification reported during execution of command according to Table 7-3
  WarningID : WORD;
  /// TRUE = overwrite an existing warning 
  Overwrite : BOOL;
END_VAR
IF ( NOT HasWarning ) OR ( Overwrite )
THEN
  THIS^.WarningID := WarningID;
END_IF
END_METHOD

END_FUNCTION_BLOCK

// Library/POUs/_internal/BaseFBs/RobotLibraryLogFB
FUNCTION_BLOCK RobotLibraryLogFB
// ------------------------------------------------------------------------- 
//  SRCI Robot Library                                                
// ------------------------------------------------------------------------- 
//                                                                           
//  Object:      RobotLibraryLogFB                                       
//  Author:      Thorsten Brach                                                
//  Date:        2024-11-10
//
//  Description:                                              
//   
//                                                                           
//  Copyright: 
//    (C) 2024 Thorsten Brach. All rights reserved                                                                                                                                            
//             Licensed under the MIT License.
//                                                                           
//  Disclaimer:                                                                           
//    This project is provided without any guarantee and can be used for   
//    private and commercial purposes. Any use is at the user’s 
//    own risk and responsibility.
//
// -------------------------------------------------------------------------
VAR_INPUT
  /// Interface to an internal logger
  InternalLogger : IMessageLogger;  
  /// Interface to an external logger
  ExternalLogger : IMessageLogger;  
  /// Logging level
  LogLevel       : LogLevelEnum := LogLevelEnum.INFO; 
END_VAR

VAR
  /// Type of the function block
 _myType         : STRING;
END_VAR

METHOD CreateLogMessage : STRING(RobotLibraryParameter.MESSAGE_TEXT_LEN)
VAR_INPUT
  /// Timestamp
  Timestamp   : SystemTime;
  /// Type of message according to Table 5-48:
  MessageType : MessageType;
  /// Severity of message according to Table 5-49: Debug, Info, Warning, Error, Fatal error
  Severity    : Severity;
  /// Code of messages
  MessageCode : DWORD;
  /// Static text of message
  MessageText : STRING(RobotLibraryParameter.MESSAGE_TEXT_LEN);  
END_VAR

VAR
  /// internal log message 
 _message    : AlarmMessage;
  /// internal string
 _tmpString  : STRING(255);
END_VAR
IF ( LogLevel <= Severity )
THEN
 _message.Timestamp   := Timestamp;
 _message.MessageType := MessageType;
 _message.Severity    := Severity;
 _message.MessageCode := MessageCode;
 _message.MessageText := StrPadRight(MyType,' ', RobotLibraryDefines.MaxTypeNameLength);
 _message.MessageText := CONCAT(_message.MessageText, ': ');
 _message.MessageText := CONCAT(_message.MessageText,MessageText);

  // return log message
  CreateLogMessage := ALARM_MESSAGE_TO_STRING(_message);
  
  // Check internal logger valid ? 
  IF ( InternalLogger <> 0 )
  THEN  
    InternalLogger.AddSystemLog( SystemLog := ALARM_MESSAGE_TO_STRING(_message));
  END_IF

  // Check external logger valid ? 
  IF ( ExternalLogger <> 0 )
  THEN  
    ExternalLogger.AddSystemLog( SystemLog := ALARM_MESSAGE_TO_STRING(_message));
  END_IF
END_IF
END_METHOD

METHOD CreateLogMessagePara1 : STRING(RobotLibraryParameter.MESSAGE_TEXT_LEN)
VAR_INPUT
  /// Timestamp
  Timestamp   : SystemTime;
  /// Type of message according to Table 5-48:
  MessageType : MessageType;
  /// Severity of message according to Table 5-49: Debug, Info, Warning, Error, Fatal error
  Severity    : Severity;
  /// Code of messages
  MessageCode : DWORD;
  /// Static text of message
  MessageText : STRING(RobotLibraryParameter.MESSAGE_TEXT_LEN);  
  /// sub string which will replace the placeholder {1}
  Para1       : STRING(RobotLibraryParameter.MESSAGE_TEXT_LEN);
END_VAR
VAR
  /// internal log message 
 _logMessage : AlarmMessage;
END_VAR
IF ( LogLevel <= Severity )
THEN
  MessageText := StrReplace(MessageText,'{1}', Para1);
  
  CreateLogMessagePara1 
    := CreateLogMessage( Timestamp   := Timestamp,
                         MessageType := MessageType,
                         Severity    := Severity,
                         MessageCode := MessageCode,
                         MessageText := MessageText);
END_IF
END_METHOD

METHOD CreateLogMessagePara2 : STRING(RobotLibraryParameter.MESSAGE_TEXT_LEN)
VAR_INPUT
  /// Timestamp
  Timestamp   : SystemTime;
  /// Type of message according to Table 5-48:
  MessageType : MessageType;
  /// Severity of message according to Table 5-49: Debug, Info, Warning, Error, Fatal error
  Severity    : Severity;
  /// Code of messages
  MessageCode : DWORD;
  /// Static text of message
  MessageText : STRING(RobotLibraryParameter.MESSAGE_TEXT_LEN);  
  /// sub string which will replace the placeholder {1}
  Para1       : STRING(RobotLibraryParameter.MESSAGE_TEXT_LEN);
  /// sub string which will replace the placeholder {2}
  Para2       : STRING(RobotLibraryParameter.MESSAGE_TEXT_LEN);
END_VAR
VAR
  /// internal log message 
 _logMessage : AlarmMessage;
END_VAR
IF ( LogLevel <= Severity )
THEN
  MessageText := StrReplace(MessageText,'{2}', Para2);
  
  CreateLogMessagePara2 
    := CreateLogMessagePara1( Timestamp   := Timestamp,
                              MessageType := MessageType,
                              Severity    := Severity,
                              MessageCode := MessageCode,
                              MessageText := MessageText,
                              Para1       := Para1);
END_IF
END_METHOD

METHOD CreateLogMessagePara3 : STRING(RobotLibraryParameter.MESSAGE_TEXT_LEN)
VAR_INPUT
  /// Timestamp
  Timestamp   : SystemTime;
  /// Type of message according to Table 5-48:
  MessageType : MessageType;
  /// Severity of message according to Table 5-49: Debug, Info, Warning, Error, Fatal error
  Severity    : Severity;
  /// Code of messages
  MessageCode : DWORD;
  /// Static text of message
  MessageText : STRING(RobotLibraryParameter.MESSAGE_TEXT_LEN);  
  /// sub string which will replace the placeholder {1}
  Para1       : STRING(RobotLibraryParameter.MESSAGE_TEXT_LEN);
  /// sub string which will replace the placeholder {2}
  Para2       : STRING(RobotLibraryParameter.MESSAGE_TEXT_LEN);
  /// sub string which will replace the placeholder {3}
  Para3       : STRING(RobotLibraryParameter.MESSAGE_TEXT_LEN);
END_VAR
VAR
  /// internal log message 
 _logMessage : AlarmMessage;
END_VAR
IF ( LogLevel <= Severity )
THEN
  MessageText := StrReplace(MessageText,'{3}', Para3);
  
  CreateLogMessagePara3
    := CreateLogMessagePara2( Timestamp   := Timestamp,
                              MessageType := MessageType,
                              Severity    := Severity,
                              MessageCode := MessageCode,
                              MessageText := MessageText,
                              Para1       := Para1,
                              Para2       := Para2);
END_IF
END_METHOD

METHOD CreateLogMessagePara4 : STRING(RobotLibraryParameter.MESSAGE_TEXT_LEN)
VAR_INPUT
  /// Timestamp
  Timestamp   : SystemTime;
  /// Type of message according to Table 5-48:
  MessageType : MessageType;
  /// Severity of message according to Table 5-49: Debug, Info, Warning, Error, Fatal error
  Severity    : Severity;
  /// Code of messages
  MessageCode : DWORD;
  /// Static text of message
  MessageText : STRING(RobotLibraryParameter.MESSAGE_TEXT_LEN);  
  /// sub string which will replace the placeholder {1}
  Para1       : STRING(RobotLibraryParameter.MESSAGE_TEXT_LEN);
  /// sub string which will replace the placeholder {2}
  Para2       : STRING(RobotLibraryParameter.MESSAGE_TEXT_LEN);
  /// sub string which will replace the placeholder {3}
  Para3       : STRING(RobotLibraryParameter.MESSAGE_TEXT_LEN);
  /// sub string which will replace the placeholder {4}
  Para4       : STRING(RobotLibraryParameter.MESSAGE_TEXT_LEN);
END_VAR
VAR
  /// internal log message 
 _logMessage : AlarmMessage;
END_VAR
IF ( LogLevel <= Severity )
THEN
  MessageText := StrReplace(MessageText,'{4}', Para4);
  
  CreateLogMessagePara4
    := CreateLogMessagePara3( Timestamp   := Timestamp,
                              MessageType := MessageType,
                              Severity    := Severity,
                              MessageCode := MessageCode,
                              MessageText := MessageText,
                              Para1       := Para1,
                              Para2       := Para2,
                              Para3       := Para3);
END_IF
END_METHOD

METHOD CreateLogMessagePara5 : STRING(RobotLibraryParameter.MESSAGE_TEXT_LEN)
VAR_INPUT
  /// Timestamp
  Timestamp   : SystemTime;
  /// Type of message according to Table 5-48:
  MessageType : MessageType;
  /// Severity of message according to Table 5-49: Debug, Info, Warning, Error, Fatal error
  Severity    : Severity;
  /// Code of messages
  MessageCode : DWORD;
  /// Static text of message
  MessageText : STRING(RobotLibraryParameter.MESSAGE_TEXT_LEN);  
  /// sub string which will replace the placeholder {1}
  Para1       : STRING(RobotLibraryParameter.MESSAGE_TEXT_LEN);
  /// sub string which will replace the placeholder {2}
  Para2       : STRING(RobotLibraryParameter.MESSAGE_TEXT_LEN);
  /// sub string which will replace the placeholder {3}
  Para3       : STRING(RobotLibraryParameter.MESSAGE_TEXT_LEN);
  /// sub string which will replace the placeholder {4}
  Para4       : STRING(RobotLibraryParameter.MESSAGE_TEXT_LEN);
  /// sub string which will replace the placeholder {5}
  Para5       : STRING(RobotLibraryParameter.MESSAGE_TEXT_LEN);
END_VAR
VAR
  /// internal log message 
 _logMessage : AlarmMessage;
END_VAR
IF ( LogLevel <= Severity )
THEN  
  MessageText := StrReplace(MessageText,'{5}', Para5);
  
  CreateLogMessagePara5
    := CreateLogMessagePara4( Timestamp   := Timestamp,
                              MessageType := MessageType,
                              Severity    := Severity,
                              MessageCode := MessageCode,
                              MessageText := MessageText,
                              Para1       := Para1,
                              Para2       := Para2,
                              Para3       := Para3,
                              Para4       := Para4);
END_IF
END_METHOD

METHOD CreateLogMessagePara6 : STRING(RobotLibraryParameter.MESSAGE_TEXT_LEN)
VAR_INPUT
  /// Timestamp
  Timestamp   : SystemTime;
  /// Type of message according to Table 5-48:
  MessageType : MessageType;
  /// Severity of message according to Table 5-49: Debug, Info, Warning, Error, Fatal error
  Severity    : Severity;
  /// Code of messages
  MessageCode : DWORD;
  /// Static text of message
  MessageText : STRING(RobotLibraryParameter.MESSAGE_TEXT_LEN);  
  /// sub string which will replace the placeholder {1}
  Para1       : STRING(RobotLibraryParameter.MESSAGE_TEXT_LEN);
  /// sub string which will replace the placeholder {2}
  Para2       : STRING(RobotLibraryParameter.MESSAGE_TEXT_LEN);
  /// sub string which will replace the placeholder {3}
  Para3       : STRING(RobotLibraryParameter.MESSAGE_TEXT_LEN);
  /// sub string which will replace the placeholder {4}
  Para4       : STRING(RobotLibraryParameter.MESSAGE_TEXT_LEN);
  /// sub string which will replace the placeholder {5}
  Para5       : STRING(RobotLibraryParameter.MESSAGE_TEXT_LEN);
  /// sub string which will replace the placeholder {6}
  Para6       : STRING(RobotLibraryParameter.MESSAGE_TEXT_LEN);
END_VAR
VAR
  /// internal log message 
 _logMessage : AlarmMessage;
END_VAR
IF ( LogLevel <= Severity )
THEN
  MessageText := StrReplace(MessageText,'{6}', Para6);
  
  CreateLogMessagePara6
    := CreateLogMessagePara5( Timestamp   := Timestamp,
                              MessageType := MessageType,
                              Severity    := Severity,
                              MessageCode := MessageCode,
                              MessageText := MessageText,
                              Para1       := Para1,
                              Para2       := Para2,
                              Para3       := Para3,
                              Para4       := Para4,
                              Para5       := Para5);
END_IF
END_METHOD

PROPERTY PROTECTED MyType : STRING
GET
MyType := _myType;
END_GET
SET
_myType := MyType;

// set the max type name length 
RobotLibraryDefines.MaxTypeNameLength := MAX(LEN(_myType), RobotLibraryDefines.MaxTypeNameLength);
END_SET
END_PROPERTY

END_FUNCTION_BLOCK

// Library/POUs/_internal/Send/RobotLibraryCommandDataFB
{attribute 'pack_mode' := '1'} 
FUNCTION_BLOCK RobotLibraryCommandDataFB EXTENDS RobotLibrarySendDataBaseFB
// ------------------------------------------------------------------------- 
//  SRCI Robot Library                                                
// ------------------------------------------------------------------------- 
//                                                                           
//  Object:      RobotLibraryCommandDataFB                                      
//  Author:      Thorsten Brach                                                
//  Date:        2025-03-29
//
//  Description:                                              
//    
//                                                                           
//  Copyright: 
//    (C) 2025 Thorsten Brach. All rights reserved                                                                                                                                            
//             Licensed under the MIT License.
//                                                                           
//  Disclaimer:                                                                           
//    This project is provided without any guarantee and can be used for   
//    private and commercial purposes. Any use is at the user’s 
//    own risk and responsibility.
//
// -------------------------------------------------------------------------

VAR_INPUT
  /// Payload
  Payload : ARRAY [0.. RobotLibraryParameter.PARAMETER_PAYLOAD_MAX] OF BYTE;
END_VAR

/// Resets the payload buffer, the payload pointer and the payload length
METHOD Reset
VAR_INPUT
END_VAR
SUPER^.Reset();

// Reset payload buffer
SysDepMemSet(pDest := ADR(Payload), Value := 0 , DataLen := SIZEOF(Payload));
END_METHOD

METHOD UpdatePointer
VAR_INPUT
END_VAR
pPayload := ADR(Payload);
END_METHOD

END_FUNCTION_BLOCK

// Library/POUs/_internal/Recv/RobotLibraryResponseDataFB
{attribute 'pack_mode' := '1'} 
FUNCTION_BLOCK RobotLibraryResponseDataFB EXTENDS RobotLibraryRecvDataBaseFB
// ------------------------------------------------------------------------- 
//  SRCI Robot Library                                                
// ------------------------------------------------------------------------- 
//                                                                           
//  Object:      RobotLibraryResponseDataFB                                       
//  Author:      Thorsten Brach                                                
//  Date:        2025-03-29
//
//  Description:                                              
//   
//                                                                           
//  Copyright: 
//    (C) 2025 Thorsten Brach. All rights reserved                                                                                                                                            
//             Licensed under the MIT License.
//                                                                           
//  Disclaimer:                                                                           
//    This project is provided without any guarantee and can be used for   
//    private and commercial purposes. Any use is at the user’s 
//    own risk and responsibility.
//
// -------------------------------------------------------------------------

VAR_INPUT
  /// Payload
  Payload    : ARRAY [0..RobotLibraryParameter.RESPONSE_PAYLOAD_MAX] OF BYTE;
END_VAR

PROPERTY IsPayloadRemaining : BOOL
GET
IsPayloadRemaining := PayloadPtr < UDINT_TO_DINT(PayloadLen );
END_GET
END_PROPERTY

/// Resets the payload buffer, the payload pointer and the payload length
METHOD Reset
VAR_INPUT
END_VAR
SUPER^.Reset();

// Reset payload buffer
SysDepMemSet(pDest := ADR(Payload), Value := 0 , DataLen := SIZEOF(Payload));
END_METHOD

METHOD UpdatePointer
VAR_INPUT
END_VAR
pPayload     := ADR(Payload);
_payloadSize := SIZEOF(Payload); // ST-FIX F22
END_METHOD

END_FUNCTION_BLOCK

// Library/POUs/_internal/Recv/RobotLibraryRecvDataBaseFB
{attribute 'pack_mode' := '1'} 
FUNCTION_BLOCK RobotLibraryRecvDataBaseFB
// ------------------------------------------------------------------------- 
//  SRCI Robot Library                                                
// ------------------------------------------------------------------------- 
//                                                                           
//  Object:      RobotLibraryRecvDataFB                                       
//  Author:      Thorsten Brach                                                
//  Date:        2024-06-01
//
//  Description:                                              
//   
//                                                                           
//  Copyright: 
//    (C) 2024 Thorsten Brach. All rights reserved                                                                                                                                            
//             Licensed under the MIT License.
//                                                                           
//  Disclaimer:                                                                           
//    This project is provided without any guarantee and can be used for   
//    private and commercial purposes. Any use is at the user’s 
//    own risk and responsibility.
//
// -------------------------------------------------------------------------
VAR_INPUT
  /// Payload length
  PayloadLen : UDINT;
  /// Payload pointer
  PayloadPtr : DINT;
END_VAR

VAR
  /// internal pointer to payload 
  pPayload : POINTER TO BYTE;
  /// Size of the payload buffer, set in UpdatePointer (ST-FIX F22)
  _payloadSize : UDINT;
END_VAR

/// returns a ArmConfigParameter from the payload buffer from the current payload pointer address and increase the payload pointer afterwards
METHOD GetArmConfig : ArmConfigParameter
VAR
  /// temporary byte
 _tmpByte : BYTE;
END_VAR
// Table 5-17: Meaning of “Config” byte
// BIT 0 Shoulder TRUE : Shoulder is Back
//                FALSE: Shoulder is Front
// BIT 1 Elbow    TRUE : Elbow is Down
//                FALSE: Elbow is Up
// BIT 2 Wrist    TRUE : Wrist is Flip
//                FALSE: Wrist is Non-Flip
// BIT 3 Spare Not used
// BIT 4 Spare Not Used
// BIT 5 Spare Not Used
// BIT 6 Spare Not Used
// BIT 7 Spare Not Used
// get 1st Byte
_tmpByte := GetByte();

IF ( _tmpByte.0 ) 
THEN
  GetArmConfig.Shoulder := ArmConfigShoulder.BACK;
ELSE
  GetArmConfig.Shoulder := ArmConfigShoulder.FRONT;
END_IF

IF ( _tmpByte.1 ) 
THEN
  GetArmConfig.Elbow := ArmConfigElbow.DOWN;
ELSE
  GetArmConfig.Elbow := ArmConfigElbow.UP;
END_IF

IF ( _tmpByte.2 ) 
THEN
  GetArmConfig.Wrist := ArmConfigWrist.FLIP;
ELSE
  GetArmConfig.Wrist := ArmConfigWrist.NON_FLIP;
END_IF


// get 2nd byte to inc the PayloadPointer
_tmpByte := GetByte();
END_METHOD

/// returns a BOOL from the payload buffer from the current payload pointer address and increase the payload pointer afterwards
METHOD GetBool : BOOL
VAR
  /// temporary byte
  _tmpByte : BYTE;
END_VAR
// update internal pointer
UpdatePointer();

// check pointer is valid ? 
IF (pPayload = RobotLibraryConstants.NULL_POINTER)
THEN
  RETURN;
END_IF


_tmpByte := GetByte();

// copy data
GetBool := _tmpByte.0;
END_METHOD

/// returns a BYTE from the payload buffer from the current payload pointer address and increase the payload pointer afterwards
METHOD GetByte : BYTE
VAR
  /// internal pointer to byte
  _tmpPointer : POINTER TO BYTE;
END_VAR
// update internal pointer
UpdatePointer();

// check pointer is valid ? 
IF (pPayload = RobotLibraryConstants.NULL_POINTER)
THEN
  RETURN;
END_IF


_tmpPointer := pPayload + DINT_TO_DWORD(PayloadPtr);

// copy data
GetByte := _tmpPointer^;
// inc payload pointer 
PayloadPtr := PayloadPtr + SIZEOF(BYTE);
END_METHOD

/// returns a datablock from the payload buffer from the current payload pointer address and increase the payload pointer afterwards
METHOD GetDataBlock
VAR_INPUT
  /// Target
  pData    : POINTER TO BYTE;
  /// Size of data block
  Size     : UDINT;
  /// Target data type is string ? 
  IsString : BOOL;
END_VAR
// update internal pointer
UpdatePointer();

// check pointer is valid ? 
IF (pPayload = RobotLibraryConstants.NULL_POINTER)
THEN
  RETURN;
END_IF


IF ( pData <> RobotLibraryConstants.NULL_POINTER)
THEN
  IF ( IsString)
  THEN
    Size := Size -1;
  END_IF

  // copy data (ST-FIX F22: only the bytes that are in the buffer, the rest is 0)
  SysDepMemSet(pDest := pData, Value := 0, DataLen := Size);
  IF ( PayloadPtr >= 0 ) AND ( DINT_TO_UDINT(PayloadPtr) < _payloadSize )
  THEN
    SysDepMemCpy(pDest   := pData,
                 pSrc    := pPayload + DINT_TO_DWORD(PayloadPtr),
                 DataLen := MIN(Size, _payloadSize - DINT_TO_UDINT(PayloadPtr)));
  END_IF
  
  // inc payload pointer 
  PayloadPtr := PayloadPtr + UDINT_TO_DINT(Size);
END_IF
END_METHOD

/// returns a DataInSync from the payload buffer from the current payload pointer address and increase the payload pointer afterwards
METHOD GetDataInSync : DataInSync
VAR
  /// temporary byte
 _tmpByte : BYTE;
END_VAR
// update internal pointer
UpdatePointer();

// check pointer is valid ? 
IF (pPayload = RobotLibraryConstants.NULL_POINTER)
THEN
  RETURN;
END_IF


// copy data
_tmpByte := GetByte();

GetDataInSync.ToolsInSync             := _tmpByte.0;
GetDataInSync.FramesInSync            := _tmpByte.1;
GetDataInSync.LoadsInSync             := _tmpByte.2;
GetDataInSync.WorkAreasInSync         := _tmpByte.3;
GetDataInSync.SoftwareLimitsInSync    := _tmpByte.4;
GetDataInSync.DefaultDynamicsInSync   := _tmpByte.5;
GetDataInSync.ReferenceDynamicsInSync := _tmpByte.6;
END_METHOD

/// returns a DWORD from the payload buffer from the current payload pointer address and increase the payload pointer afterwards
METHOD GetDword : DWORD
// update internal pointer
UpdatePointer();

// check pointer is valid ? 
IF (pPayload = RobotLibraryConstants.NULL_POINTER)
THEN
  RETURN;
END_IF

// copy data
SysDepMemCpy(pDest := ADR(GetDword), pSrc := pPayload + DINT_TO_DWORD(PayloadPtr), DataLen := SIZEOF(DWORD));
// inc payload pointer 
PayloadPtr := PayloadPtr + SIZEOF(DWORD);
END_METHOD

/// returns a FragmentAction from the payload buffer from the current payload pointer address and increase the payload pointer afterwards
METHOD GetFragmentAction : FragmentAction
VAR
  /// temporary byte
 _tmpByte : BYTE;
END_VAR
// update internal pointer
UpdatePointer();

// check pointer is valid ? 
IF (pPayload = RobotLibraryConstants.NULL_POINTER)
THEN
  RETURN;
END_IF

// copy data
_tmpByte := GetByte();

GetFragmentAction.Complete := _tmpByte.0;
GetFragmentAction.Reset    := _tmpByte.1;
GetFragmentAction.Clear    := _tmpByte.2;
GetFragmentAction.BIT03    := _tmpByte.3;
GetFragmentAction.BIT04    := _tmpByte.4;
GetFragmentAction.BIT05    := _tmpByte.5;
GetFragmentAction.BIT06    := _tmpByte.6;
GetFragmentAction.BIT07    := _tmpByte.7;
END_METHOD

/// returns the 1st halfe BYTE from the payload buffer from the current payload pointer address and increase the payload pointer afterwards
METHOD GetHalfeByte1 : BYTE
VAR_INPUT
  /// Increase payload pointer 
  IncPayloadPtr : BOOL;
END_VAR

VAR
  /// temporary byte
 _tmpByte    : BYTE;
  /// internal pointer to byte
 _tmpPointer : POINTER TO BYTE;
END_VAR
// update internal pointer
UpdatePointer();

// check pointer is valid ? 
IF (pPayload = RobotLibraryConstants.NULL_POINTER)
THEN
  RETURN;
END_IF

// set pointer
_tmpPointer := pPayload + DINT_TO_DWORD(PayloadPtr); 
// copy data
_tmpByte := _tmpPointer^;

GetHalfeByte1.0 := _tmpByte.0;
GetHalfeByte1.1 := _tmpByte.1;
GetHalfeByte1.2 := _tmpByte.2;
GetHalfeByte1.3 := _tmpByte.3;

IF (IncPayloadPtr)
THEN  
  // inc payload pointer
  PayloadPtr := PayloadPtr + SIZEOF(BYTE);
END_IF
END_METHOD

/// returns the 1st halfe BYTE from the payload buffer from the current payload pointer address and increase the payload pointer afterwards
METHOD GetHalfeByte2 : BYTE
VAR_INPUT
  /// Increase payload pointer 
  IncPayloadPtr : BOOL;
END_VAR

VAR
  /// temporary byte
 _tmpByte    : BYTE;
  /// internal pointer to byte
 _tmpPointer : POINTER TO BYTE;
END_VAR
// update internal pointer
UpdatePointer();

// check pointer is valid ? 
IF (pPayload = RobotLibraryConstants.NULL_POINTER)
THEN
  RETURN;
END_IF

// set pointer
_tmpPointer := pPayload + DINT_TO_DWORD(PayloadPtr); 
// copy data
_tmpByte := _tmpPointer^;

GetHalfeByte2.0 := _tmpByte.4;
GetHalfeByte2.1 := _tmpByte.5;
GetHalfeByte2.2 := _tmpByte.6;
GetHalfeByte2.3 := _tmpByte.7;

IF (IncPayloadPtr)
THEN  
  // inc payload pointer
  PayloadPtr := PayloadPtr + SIZEOF(BYTE);
END_IF
END_METHOD

/// returns a IEC_Date from the payload buffer from the current payload pointer address and increase the payload pointer afterwards
METHOD GetIecDate : IEC_Date
// update internal pointer
UpdatePointer();

// check pointer is valid ? 
IF (pPayload = RobotLibraryConstants.NULL_POINTER)
THEN
  RETURN;
END_IF

// copy data
SysDepMemCpy(pDest := ADR(GetIecDate), pSrc := pPayload + DINT_TO_DWORD(PayloadPtr), DataLen := SIZEOF(IEC_DATE));
// swap byte order
GetIecDate := SwapIecDate(GetIecDate);
// inc payload pointer   
PayloadPtr := PayloadPtr + SIZEOF(IEC_DATE);
END_METHOD

/// returns a IEC_TIME from the payload buffer from the current payload pointer address and increase the payload pointer afterwards
METHOD GetIecTime : IEC_TIME
// update internal pointer
UpdatePointer();

// check pointer is valid ? 
IF (pPayload = RobotLibraryConstants.NULL_POINTER)
THEN
  RETURN;
END_IF

// copy data
SysDepMemCpy(pDest := ADR(GetIecTime), pSrc := pPayload + DINT_TO_DWORD(PayloadPtr), DataLen := SIZEOF(IEC_TIME));
// swap byte order
GetIecTime := SwapIecTime(GetIecTime);
// inc payload pointer   
PayloadPtr := PayloadPtr + SIZEOF(IEC_TIME);
END_METHOD

/// returns a INT from the payload buffer from the current payload pointer address and increase the payload pointer afterwards
METHOD GetInt : INT
// update internal pointer
UpdatePointer();

// check pointer is valid ? 
IF (pPayload = RobotLibraryConstants.NULL_POINTER)
THEN
  RETURN;
END_IF

// copy data
SysDepMemCpy(pDest := ADR(GetInt), pSrc := pPayload + DINT_TO_DWORD(PayloadPtr), DataLen := SIZEOF(INT));
// swap byte order
GetInt := SwapInt(GetInt);
// inc payload pointer   
PayloadPtr := PayloadPtr + SIZEOF(INT);
END_METHOD

/// returns a REAL from the payload buffer from the current payload pointer address and increase the payload pointer afterwards
METHOD GetReal : REAL
// update internal pointer
UpdatePointer();

// check pointer is valid ? 
IF (pPayload = RobotLibraryConstants.NULL_POINTER)
THEN
  RETURN;
END_IF

// copy data
SysDepMemCpy(pDest := ADR(GetReal), pSrc := pPayload + DINT_TO_DWORD(PayloadPtr), DataLen := SIZEOF(REAL));
// swap byte order
GetReal := SwapReal(GetReal);
// inc payload pointer   
PayloadPtr := PayloadPtr + SIZEOF(Real);
END_METHOD

/// returns a SINT from the payload buffer from the current payload pointer address and increase the payload pointer afterwards
METHOD GetSint : SINT
// update internal pointer
UpdatePointer();

// check pointer is valid ? 
IF (pPayload = RobotLibraryConstants.NULL_POINTER)
THEN
  RETURN;
END_IF

// copy data
SysDepMemCpy(pDest := ADR(GetSint), pSrc := pPayload + DINT_TO_DWORD(PayloadPtr), DataLen := SIZEOF(SINT));
// inc payload pointer 
PayloadPtr := PayloadPtr + SIZEOF(SINT);
END_METHOD

/// returns a String from the payload buffer from the current payload pointer address and increase the payload pointer afterwards
METHOD GetString : STRING(255)
VAR_INPUT
  Size : DINT;
END_VAR
// update internal pointer
UpdatePointer();

// check pointer is valid ? 
IF (pPayload = RobotLibraryConstants.NULL_POINTER)
THEN
  RETURN;
END_IF

// copy data
SysDepMemCpy(pDest := ADR(GetString), pSrc := pPayload + DINT_TO_DWORD(PayloadPtr), DataLen := DINT_TO_UDINT(Size));

// inc payload pointer 
PayloadPtr := PayloadPtr + Size;
END_METHOD

/// returns a TrackingStatus from the payload buffer from the current payload pointer address and increase the payload pointer afterwards
METHOD GetTrackingStatus : TrackingStatus
VAR
  /// temporary byte
  tmpByte : BYTE;
END_VAR
// update internal pointer
UpdatePointer();

// check pointer is valid ? 
IF (pPayload = RobotLibraryConstants.NULL_POINTER)
THEN
  RETURN;
END_IF

// copy data
tmpByte := GetByte();

GetTrackingStatus.ConveyorTrackingEnabled   := tmpByte.0;  
GetTrackingStatus.WaitingForSynchronization := tmpByte.1;
GetTrackingStatus.Synchronizing             := tmpByte.2;
GetTrackingStatus.Synchronous               := tmpByte.3;
GetTrackingStatus.Desynchronizing           := tmpByte.4;
GetTrackingStatus.SyncOutZoneEntered        := tmpByte.5;
GetTrackingStatus.SyncOutZoneLeft           := tmpByte.6;
GetTrackingStatus.NotUsed                   := tmpByte.7;
END_METHOD

/// returns a TurnNumber from the payload buffer from the current payload pointer address and increase the payload pointer afterwards
METHOD GetTurnNumbers : TurnNumber
// update internal pointer
UpdatePointer();

// check pointer is valid ? 
IF (pPayload = RobotLibraryConstants.NULL_POINTER)
THEN
  RETURN;
END_IF

GetTurnNumbers.J1Turns := SIGN_MAGNITUDE_TO_TURN(Value := GetHalfeByte1(FALSE), Bits := 3); // ST-FIX F3
GetTurnNumbers.J2Turns := SIGN_MAGNITUDE_TO_TURN(Value := GetHalfeByte2(TRUE),  Bits := 3); // ST-FIX F3

GetTurnNumbers.J3Turns := SIGN_MAGNITUDE_TO_TURN(Value := GetHalfeByte1(FALSE), Bits := 3); // ST-FIX F3
GetTurnNumbers.J4Turns := SIGN_MAGNITUDE_TO_TURN(Value := GetHalfeByte2(TRUE),  Bits := 3); // ST-FIX F3

GetTurnNumbers.J5Turns := SIGN_MAGNITUDE_TO_TURN(Value := GetHalfeByte1(FALSE), Bits := 3); // ST-FIX F3
GetTurnNumbers.J6Turns := SIGN_MAGNITUDE_TO_TURN(Value := GetHalfeByte2(TRUE),  Bits := 3); // ST-FIX F3

GetTurnNumbers.E1Turns := SIGN_MAGNITUDE_TO_TURN(Value := GetByte(), Bits := 7); // ST-FIX F3
END_METHOD

/// returns a UDINT from the payload buffer from the current payload pointer address and increase the payload pointer afterwards
METHOD GetUdint : UDINT
// update internal pointer
UpdatePointer();

// check pointer is valid ? 
IF (pPayload = RobotLibraryConstants.NULL_POINTER)
THEN
  RETURN;
END_IF

// copy data
SysDepMemCpy(pDest := ADR(GetUdint), pSrc := pPayload + DINT_TO_DWORD(PayloadPtr), DataLen := SIZEOF(UDINT));
// swap byte order
GetUdint := SwapUdint(GetUdint);
// inc payload pointer   
PayloadPtr := PayloadPtr + SIZEOF(UDINT);
END_METHOD

/// returns a UINT from the payload buffer from the current payload pointer address and increase the payload pointer afterwards
METHOD GetUint : UINT
// update internal pointer
UpdatePointer();

// check pointer is valid ? 
IF (pPayload = RobotLibraryConstants.NULL_POINTER)
THEN
  RETURN;
END_IF

// copy data
SysDepMemCpy(pDest := ADR(GetUint), pSrc := pPayload + DINT_TO_DWORD(PayloadPtr), DataLen := SIZEOF(UINT));
// swap byte order
GetUint := SwapUint(GetUint);
// inc payload pointer   
PayloadPtr := PayloadPtr + SIZEOF(UINT);
END_METHOD

/// returns a USINT from the payload buffer from the current payload pointer address and increase the payload pointer afterwards
METHOD GetUsint : USINT
// update internal pointer
UpdatePointer();

// check pointer is valid ? 
IF (pPayload = RobotLibraryConstants.NULL_POINTER)
THEN
  RETURN;
END_IF

// copy data
SysDepMemCpy(pDest := ADR(GetUsint), pSrc := pPayload + DINT_TO_DWORD(PayloadPtr), DataLen := SIZEOF(USINT));
// inc payload pointer 
PayloadPtr := PayloadPtr + SIZEOF(USINT);
END_METHOD

/// returns a WORD from the payload buffer from the current payload pointer address and increase the payload pointer afterwards
METHOD GetWord : WORD
// update internal pointer
UpdatePointer();

// check pointer is valid ? 
IF (pPayload = RobotLibraryConstants.NULL_POINTER)
THEN
  RETURN;
END_IF

// copy data
SysDepMemCpy(pDest := ADR(GetWord), pSrc := pPayload + DINT_TO_DWORD(PayloadPtr), DataLen := SIZEOF(WORD));
// swap byte order
GetWord := SwapWord(GetWord);
// inc payload pointer   
PayloadPtr := PayloadPtr + SIZEOF(WORD);
END_METHOD

/// Resets the payload buffer, the payload pointer and the payload length
METHOD Reset
VAR_INPUT
END_VAR
PayloadLen := 0;
PayloadPtr := 0;
END_METHOD

METHOD UpdatePointer
VAR_INPUT
END_VAR
END_METHOD

END_FUNCTION_BLOCK

// Library/POUs/_internal/Recv/RobotLibraryRecvDataFB
{attribute 'pack_mode' := '1'} 
FUNCTION_BLOCK RobotLibraryRecvDataFB EXTENDS RobotLibraryRecvDataBaseFB
// ------------------------------------------------------------------------- 
//  SRCI Robot Library                                                
// ------------------------------------------------------------------------- 
//                                                                           
//  Object:      RobotLibraryRecvDataFB                                       
//  Author:      Thorsten Brach                                                
//  Date:        2024-06-01
//
//  Description:                                              
//   
//                                                                           
//  Copyright: 
//    (C) 2024 Thorsten Brach. All rights reserved                                                                                                                                            
//             Licensed under the MIT License.
//                                                                           
//  Disclaimer:                                                                           
//    This project is provided without any guarantee and can be used for   
//    private and commercial purposes. Any use is at the user’s 
//    own risk and responsibility.
//
// -------------------------------------------------------------------------
VAR_INPUT
  /// Payload
  Payload    : POINTER TO BYTE;
  /// Size of the Payload array
  PayLoadSize : UDINT;
END_VAR

METHOD GetLifeSignFooter : BYTE
VAR
  /// temporary 
  pLifeSign : POINTER TO BYTE;
END_VAR
pLifeSign := Payload + PayLoadSize -1;


GetLifeSignFooter := GetHalfeByteHi(pLifeSign^);
END_METHOD

METHOD UpdatePointer
VAR_INPUT
END_VAR
pPayload     := Payload;
_payloadSize := PayLoadSize; // ST-FIX F22
END_METHOD

END_FUNCTION_BLOCK

// Library/POUs/Additional/MC_ExchangeConfiguration/MC_ExchangeConfigurationFB
/// Reads and writes specific configuration parameters on RC that are required for the RI to work
FUNCTION_BLOCK MC_ExchangeConfigurationFB EXTENDS RobotLibraryBaseEnableFB
// ------------------------------------------------------------------------- 
//  SRCI Robot Library                                                
// ------------------------------------------------------------------------- 
//                                                                           
//  Object:      ExchangeConfigurationFB                                       
//  Author:      Thorsten Brach                                                
//  Date:        2024-06-01
//
//  Description:                                              
//   
//                                                                           
//  Copyright: 
//    (C) 2024 Thorsten Brach. All rights reserved                                                                                                                                            
//             Licensed under the MIT License.
//                                                                           
//  Disclaimer:                                                                           
//    This project is provided without any guarantee and can be used for   
//    private and commercial purposes. Any use is at the user’s 
//    own risk and responsibility.
//
// -------------------------------------------------------------------------
VAR_INPUT
  /// Command parameter 
  ParCmd            : ExchangeConfigurationParCmd;
END_VAR

VAR_OUTPUT
  /// Command is transferred and confirmed by the RC
  CommandBuffered   : BOOL;
  /// Receiving of input parameter values has been acknowledged by RC
  ParameterAccepted : BOOL;
  /// command results
  OutCmd            : ExchangeConfigurationOutCmd;
END_VAR

VAR
  /// internal copy of command parameter 
 _parCmd            : ExchangeConfigurationParCmd;
  /// command data to send
 _command           : ExchangeConfigurationSendData;
  /// response data received
 _response          : ExchangeConfigurationRecvData;
END_VAR

SUPER^(AxesGroup := AxesGroup);

METHOD INTERNAL CheckAddParameter : BOOL
VAR_INPUT
  /// Payload pointer
  PayloadPtr : UDINT;
END_VAR
VAR
  /// Payload as byte array
  Payload    : ARRAY [1..SIZEOF(_command)] OF BYTE;
  /// Null Byte array 
  Null       : ARRAY [1..SIZEOF(_command)] OF BYTE;
  /// Data length to compare
  DataLen    : UDINT;
END_VAR
// Payload pointer must be decreased by one byte, because ADR(Payload) is already one byte !
PayloadPtr := LIMIT (0, PayloadPtr - 1, SIZEOF(Payload) -1);
// Convert command struct to payload array
SysDepMemCpy( pDest := ADR(Payload), pSrc := ADR(_command), DataLen := SIZEOF(_command));
// Calculate the data length to compare - at least one byte must be compared !
DataLen := LIMIT(1, SIZEOF(Payload) - PayloadPtr, SIZEOF(Payload)); 
// Compare Payload-Array with Null-Byte-Array
CheckAddParameter := SysDepMemCmp( pData1 := ADR(Payload) + PayloadPtr , pData2 := ADR(Null), DataLen := DataLen) <>  RobotLibraryConstants.OK ;
END_METHOD

METHOD PROTECTED CheckFunctionSupported : BOOL
VAR_IN_OUT
  /// Robot assignment of function
  AxesGroup : AxesGroup; 
END_VAR
CheckFunctionSupported := TRUE; // Function is mandatory 
RETURN;

CheckFunctionSupported := AxesGroup.State.RobotData.RCSupportedFunctions.ExchangeConfiguration;

IF ( NOT CheckFunctionSupported )
THEN
  // call base implementation for set error and create log entry
  SUPER^.CheckFunctionSupported(AxesGroup := AxesGroup);
END_IF
END_METHOD

METHOD PROTECTED CheckParameterChanged : BOOL
VAR_IN_OUT
  /// Robot assignment of function
  AxesGroup    : AxesGroup; 
END_VAR
// Check ParCmd Size is > 0, because MemCmp does not work correctly with size = 0
IF (SIZEOF(ParCmd) = 0) OR (_stepCmd = 0)
THEN 
  RETURN;
END_IF

// compare memory 
_parameterChanged := ( SysDepMemCmp(pData1 := ADR(ParCmd), pData2 := ADR(_parCmd), DataLen := SIZEOF(ParCmd)) <> RobotLibraryConstants.OK );

// check parameter valid ?
_parameterValid   := CheckParameterValid( AxesGroup := AxesGroup );

IF ((  _parameterChanged        )  AND 
    (  _parameterValid          )) OR
    (  _parameterUpdateInternal )  
THEN  
  // Create log entry for parameter changed event
  CreateLogMessagePara1 ( Timestamp   := AxesGroup.State.SystemTime,
                          MessageType := MessageType.CMD,
                          Severity    := Severity.DEBUG,
                          MessageCode := 0,
                          MessageText := 'NotifyParameterChanged Event {1}',
                          Para1       :=  '' );

  // reset internal flag for send parameter update
 _parameterUpdateInternal := FALSE;
  // update internal copy of parameters 
 _parCmd := ParCmd;
  // inc parameter sequence
 _command.ParSeq := _command.ParSeq + 1;
  // update command data  
  CommandData := CreateCommandPayload(AxesGroup := AxesGroup); // ( Access via reference to rCommandFB in ACR )
  // notify active command register 
  AxesGroup.Acyclic.ActiveCommandRegister.NotifyParameterChanged := _uniqueID;
  // Reset parameter accepted flag
  ParameterAccepted := FALSE;
END_IF
END_METHOD

METHOD PROTECTED CheckParameterValid : BOOL
VAR_IN_OUT
  /// Robot assignment of function
  AxesGroup : AxesGroup; 
END_VAR
CheckParameterValid := TRUE;

// Check ParCmd.LogLevel valid ? 
IF (( ParCmd.LogLevel <> Severity.DEACTIVATE  ) AND  
    ( ParCmd.LogLevel <> Severity.DEBUG       ) AND
    ( ParCmd.LogLevel <> Severity.INFO        ) AND
    ( ParCmd.LogLevel <> Severity.WARNING     ) AND
    ( ParCmd.LogLevel <> Severity.ERROR       ) AND
    ( ParCmd.LogLevel <> Severity.FATAL_ERROR ))    
THEN
  // Parameter not valid
  CheckParameterValid := FALSE;
  // Set error
  SetError( ErrorID := RobotLibraryErrorIdEnum.ERR_INVALID_PAR_CMD, Overwrite := TRUE );
  // Create log entry
  CreateLogMessagePara1 ( Timestamp   := AxesGroup.State.SystemTime,
                          MessageType := MessageType.CMD,
                          Severity    := Severity.ERROR,
                          MessageCode := ErrorID,
                          MessageText := 'Invalid Parameter ParCmd.LogLevel = {1}',
                          Para1       :=  LOG_LEVEL_TO_STRING(ParCmd.LogLevel));
  RETURN;                          
END_IF


// Check ParCmd.WaitAtBlendingZone
// -> no plausibility check for boolean


// Check ParCmd.AllowSecSeqWhileSubprogram
// -> no plausibility check for boolean


// Check ParCmd.DelayTime valid ? 
IF ( ParCmd.DelayTime < 0  )   
THEN
  // Parameter not valid
  CheckParameterValid := FALSE;
  // Set error
  SetError( ErrorID := RobotLibraryErrorIdEnum.ERR_INVALID_PAR_CMD, Overwrite := TRUE );
  // Create log entry
  CreateLogMessagePara1 ( Timestamp   := AxesGroup.State.SystemTime,
                          MessageType := MessageType.CMD,
                          Severity    := Severity.ERROR,
                          MessageCode := ErrorID,
                          MessageText := 'Invalid Parameter ParCmd.DelayTime = {1} ms',
                          Para1       :=  UINT_TO_STRING(ParCmd.DelayTime));
  RETURN;                          
END_IF


// Check ParCmd.WaitForNrOfCmd valid ? 
IF ( ParCmd.WaitForNrOfCmd < 0  )   
THEN
  // Parameter not valid
  CheckParameterValid := FALSE;
  // Set error
  SetError( ErrorID := RobotLibraryErrorIdEnum.ERR_INVALID_PAR_CMD , Overwrite :=  TRUE );
  // Create log entry
  CreateLogMessagePara1 ( Timestamp   := AxesGroup.State.SystemTime,
                          MessageType := MessageType.CMD,
                          Severity    := Severity.ERROR,
                          MessageCode := ErrorID,
                          MessageText := 'Invalid Parameter ParCmd.WaitForNrOfCmd = {1}',
                          Para1       :=  UINT_TO_STRING(ParCmd.WaitForNrOfCmd));
  RETURN;                          
END_IF


// Check ParCmd.LifeSignTimeOut valid ? 
IF ( ParCmd.LifeSignTimeOut < 10 )   
THEN
  // Parameter not valid
  CheckParameterValid := FALSE;
  // Set error
  SetError( ErrorID := RobotLibraryErrorIdEnum.ERR_INVALID_PAR_CMD, Overwrite := TRUE );
  // Create log entry
  CreateLogMessagePara1 ( Timestamp   := AxesGroup.State.SystemTime,
                          MessageType := MessageType.CMD,
                          Severity    := Severity.ERROR,
                          MessageCode := ErrorID,
                          MessageText := 'Invalid Parameter ParCmd.LifeSignTimeOut = {1} ms',
                          Para1       :=  UINT_TO_STRING(ParCmd.LifeSignTimeOut));
  RETURN;                          
END_IF


